Universal Robots URScript: FaiChun_9 Jan_1.script

def Machining1():
  # Default parameters:
  global speed_ms = 0.01
  global speed_rads = 0.75
  global accel_mss = 3
  global accel_radss = 1.2
  global blend_radius_m = 0.0003

  # Add subprograms here
  # Start of main program
  # Program generated by RoboDK v5.6.8 for UR10e on 09/01/2025 14:53:28
  # Using nominal kinematics.
  blend_radius_m = 0.0003
  speed_ms = 0.01
  # set_reference(p[0.305000, -0.155000, 0.000000, 0.000000, 0.000000, 0.000000])
  set_tcp(p[0.000000, 0.000000, 0.252000, 0.000000, 0.000000, 0.000000])
  # Show Tool
  movej([0.378214, -1.028418, -2.649277, -1.034694, 1.570796, 1.949010],accel_radss,speed_rads,0,blend_radius_m)
  movel([0.378214, -1.088062, -2.690368, -0.933959, 1.570796, 1.949010],accel_mss,speed_ms,0,blend_radius_m)
  #SetTool1
  #M_RunCode6
  #SetRPM60000
  speed_ms = 0.01
  #M_RunCode3
  movel([0.378214, -1.116012, -2.706101, -0.890276, 1.570796, 1.949010],accel_mss,speed_ms,0,blend_radius_m)
  speed_ms = 0.003
  movel([0.378214, -1.123422, -2.709978, -0.878989, 1.570796, 1.949010],accel_mss,speed_ms,0,blend_radius_m)
  speed_ms = 0.007
  movel([0.427669, -1.206915, -2.673266, -0.832208, 1.570796, 1.998465],accel_mss,speed_ms,0,blend_radius_m)
  movel([0.418964, -1.213811, -2.669903, -0.828675, 1.570796, 1.989761],accel_mss,speed_ms,0,blend_radius_m)
  movel([0.421470, -1.218334, -2.667668, -0.826387, 1.570796, 1.992267],accel_mss,speed_ms,0,blend_radius_m)
  movel([0.423710, -1.216572, -2.668541, -0.827276, 1.570796, 1.994506],accel_mss,speed_ms,0,blend_radius_m)
  movel([0.422070, -1.213581, -2.670016, -0.828792, 1.570796, 1.992867],accel_mss,speed_ms,0,blend_radius_m)
  movel([0.428515, -1.208497, -2.672499, -0.831392, 1.570796, 1.999312],accel_mss,speed_ms,0,blend_radius_m)
  movel([0.428905, -1.209227, -2.672145, -0.831017, 1.570796, 1.999701],accel_mss,speed_ms,0,blend_radius_m)
  movel([0.430913, -1.212978, -2.670312, -0.829099, 1.570796, 2.001710],accel_mss,speed_ms,0,blend_radius_m)
  movel([0.426574, -1.216377, -2.668637, -0.827374, 1.570796, 1.997371],accel_mss,speed_ms,0,blend_radius_m)
  movel([0.427415, -1.217932, -2.667867, -0.826590, 1.570796, 1.998211],accel_mss,speed_ms,0,blend_radius_m)
  movel([0.431749, -1.214549, -2.669539, -0.828300, 1.570796, 2.002545],accel_mss,speed_ms,0,blend_radius_m)
  movel([0.434110, -1.219016, -2.667329, -0.826045, 1.570796, 2.004906],accel_mss,speed_ms,0,blend_radius_m)
  movel([0.429796, -1.222362, -2.665657, -0.824369, 1.570796, 2.000592],accel_mss,speed_ms,0,blend_radius_m)
  movel([0.431384, -1.225346, -2.664156, -0.822886, 1.570796, 2.002180],accel_mss,speed_ms,0,blend_radius_m)
  movel([0.425058, -1.230240, -2.661672, -0.820476, 1.570796, 1.995855],accel_mss,speed_ms,0,blend_radius_m)
  movel([0.423449, -1.227294, -2.663171, -0.821924, 1.570796, 1.994246],accel_mss,speed_ms,0,blend_radius_m)
  movel([0.421238, -1.229018, -2.662295, -0.821076, 1.570796, 1.992034],accel_mss,speed_ms,0,blend_radius_m)
  movel([0.422852, -1.231953, -2.660796, -0.819639, 1.570796, 1.993648],accel_mss,speed_ms,0,blend_radius_m)
  movel([0.417606, -1.236027, -2.658699, -0.817662, 1.570796, 1.988403],accel_mss,speed_ms,0,blend_radius_m)
  movel([0.416595, -1.236817, -2.658291, -0.817282, 1.570796, 1.987391],accel_mss,speed_ms,0,blend_radius_m)
  movel([0.414170, -1.232527, -2.660502, -0.819360, 1.570796, 1.984966],accel_mss,speed_ms,0,blend_radius_m)
  movel([0.418408, -1.229206, -2.662200, -0.820984, 1.570796, 1.989204],accel_mss,speed_ms,0,blend_radius_m)
  movel([0.417558, -1.227687, -2.662972, -0.821730, 1.570796, 1.988355],accel_mss,speed_ms,0,blend_radius_m)
  movel([0.411120, -1.232746, -2.660390, -0.819253, 1.570796, 1.981917],accel_mss,speed_ms,0,blend_radius_m)
  movel([0.414410, -1.238516, -2.657409, -0.816464, 1.570796, 1.985206],accel_mss,speed_ms,0,blend_radius_m)
  movel([0.308742, -1.323345, -2.608871, -0.780173, 1.570796, 1.879539],accel_mss,speed_ms,0,blend_radius_m)
  movel([0.217512, -1.401117, -2.555954, -0.755318, 1.570796, 1.788308],accel_mss,speed_ms,0,blend_radius_m)
  movel([0.213488, -1.397361, -2.558708, -0.756321, 1.570796, 1.784284],accel_mss,speed_ms,0,blend_radius_m)
  movel([0.208744, -1.401573, -2.555618, -0.755198, 1.570796, 1.779541],accel_mss,speed_ms,0,blend_radius_m)
  movel([0.209793, -1.402537, -2.554907, -0.754944, 1.570796, 1.780589],accel_mss,speed_ms,0,blend_radius_m)
  movel([0.212909, -1.399774, -2.556941, -0.755674, 1.570796, 1.783706],accel_mss,speed_ms,0,blend_radius_m)
  movel([0.215882, -1.402546, -2.554901, -0.754942, 1.570796, 1.786679],accel_mss,speed_ms,0,blend_radius_m)
  movel([0.215131, -1.403208, -2.554412, -0.754769, 1.570796, 1.785928],accel_mss,speed_ms,0,blend_radius_m)
  movel([0.211277, -1.406609, -2.551890, -0.753890, 1.570796, 1.782073],accel_mss,speed_ms,0,blend_radius_m)
  movel([0.209269, -1.404754, -2.553268, -0.754367, 1.570796, 1.780066],accel_mss,speed_ms,0,blend_radius_m)
  movel([0.207663, -1.406180, -2.552209, -0.754000, 1.570796, 1.778459],accel_mss,speed_ms,0,blend_radius_m)
  movel([0.209672, -1.408029, -2.550833, -0.753528, 1.570796, 1.780468],accel_mss,speed_ms,0,blend_radius_m)
  movel([0.205118, -1.412065, -2.547809, -0.752515, 1.570796, 1.775914],accel_mss,speed_ms,0,blend_radius_m)
  movel([0.203102, -1.410238, -2.549181, -0.752970, 1.570796, 1.773898],accel_mss,speed_ms,0,blend_radius_m)
  movel([0.200044, -1.412967, -2.547130, -0.752292, 1.570796, 1.770840],accel_mss,speed_ms,0,blend_radius_m)
  movel([0.197039, -1.410284, -2.549146, -0.752959, 1.570796, 1.767835],accel_mss,speed_ms,0,blend_radius_m)
  movel([0.200101, -1.407535, -2.551201, -0.753653, 1.570796, 1.770897],accel_mss,speed_ms,0,blend_radius_m)
  movel([0.199043, -1.406589, -2.551905, -0.753895, 1.570796, 1.769840],accel_mss,speed_ms,0,blend_radius_m)
  movel([0.195980, -1.409343, -2.549851, -0.753195, 1.570796, 1.766776],accel_mss,speed_ms,0,blend_radius_m)
  movel([0.193434, -1.407104, -2.551522, -0.753763, 1.570796, 1.764230],accel_mss,speed_ms,0,blend_radius_m)
  movel([0.192941, -1.406669, -2.551845, -0.753874, 1.570796, 1.763737],accel_mss,speed_ms,0,blend_radius_m)
  movel([0.197491, -1.402558, -2.554892, -0.754939, 1.570796, 1.768287],accel_mss,speed_ms,0,blend_radius_m)
  movel([0.199540, -1.404383, -2.553543, -0.754463, 1.570796, 1.770337],accel_mss,speed_ms,0,blend_radius_m)
  movel([0.201142, -1.402944, -2.554607, -0.754838, 1.570796, 1.771938],accel_mss,speed_ms,0,blend_radius_m)
  movel([0.198026, -1.400161, -2.556657, -0.755571, 1.570796, 1.768823],accel_mss,speed_ms,0,blend_radius_m)
  movel([0.191871, -1.405733, -2.552541, -0.754115, 1.570796, 1.762667],accel_mss,speed_ms,0,blend_radius_m)
  movel([0.191373, -1.405301, -2.552862, -0.754226, 1.570796, 1.762169],accel_mss,speed_ms,0,blend_radius_m)
  movel([0.131815, -1.358213, -2.586196, -0.767981, 1.570796, 1.702611],accel_mss,speed_ms,0,blend_radius_m)
  movel([0.062823, -1.314529, -2.614344, -0.783517, 1.570796, 1.633619],accel_mss,speed_ms,0,blend_radius_m)
  movel([0.069044, -1.307429, -2.618676, -0.786284, 1.570796, 1.639841],accel_mss,speed_ms,0,blend_radius_m)
  movel([0.064886, -1.305093, -2.620087, -0.787209, 1.570796, 1.635683],accel_mss,speed_ms,0,blend_radius_m)
  movel([0.063265, -1.306951, -2.618965, -0.786472, 1.570796, 1.634061],accel_mss,speed_ms,0,blend_radius_m)
  movel([0.066004, -1.308479, -2.618039, -0.785870, 1.570796, 1.636801],accel_mss,speed_ms,0,blend_radius_m)
  movel([0.061405, -1.313734, -2.614831, -0.783823, 1.570796, 1.632201],accel_mss,speed_ms,0,blend_radius_m)
  movel([0.060750, -1.313370, -2.615055, -0.783964, 1.570796, 1.631546],accel_mss,speed_ms,0,blend_radius_m)
  movel([0.057348, -1.311503, -2.616198, -0.784688, 1.570796, 1.628144],accel_mss,speed_ms,0,blend_radius_m)
  movel([0.060443, -1.307941, -2.618366, -0.786082, 1.570796, 1.631240],accel_mss,speed_ms,0,blend_radius_m)
  movel([0.059013, -1.307156, -2.618841, -0.786392, 1.570796, 1.629809],accel_mss,speed_ms,0,blend_radius_m)
  movel([0.055918, -1.310726, -2.616672, -0.784991, 1.570796, 1.626714],accel_mss,speed_ms,0,blend_radius_m)
  movel([0.051821, -1.308523, -2.618013, -0.785853, 1.570796, 1.622617],accel_mss,speed_ms,0,blend_radius_m)
  movel([0.054912, -1.304932, -2.620184, -0.787273, 1.570796, 1.625709],accel_mss,speed_ms,0,blend_radius_m)
  movel([0.052126, -1.303438, -2.621082, -0.787868, 1.570796, 1.622923],accel_mss,speed_ms,0,blend_radius_m)
  movel([0.056741, -1.298064, -2.624290, -0.790035, 1.570796, 1.627538],accel_mss,speed_ms,0,blend_radius_m)
  movel([0.059531, -1.299576, -2.623391, -0.789421, 1.570796, 1.630327],accel_mss,speed_ms,0,blend_radius_m)
  movel([0.061161, -1.297689, -2.624513, -0.790187, 1.570796, 1.631957],accel_mss,speed_ms,0,blend_radius_m)
  movel([0.058371, -1.296169, -2.625412, -0.790807, 1.570796, 1.629167],accel_mss,speed_ms,0,blend_radius_m)
  movel([0.062287, -1.291620, -2.628088, -0.792681, 1.570796, 1.633084],accel_mss,speed_ms,0,blend_radius_m)
  movel([0.063052, -1.290735, -2.628605, -0.793049, 1.570796, 1.633848],accel_mss,speed_ms,0,blend_radius_m)
  movel([0.067186, -1.293020, -2.627267, -0.792102, 1.570796, 1.637983],accel_mss,speed_ms,0,blend_radius_m)
  movel([0.064017, -1.296673, -2.625115, -0.790602, 1.570796, 1.634813],accel_mss,speed_ms,0,blend_radius_m)
  movel([0.065457, -1.297471, -2.624642, -0.790276, 1.570796, 1.636253],accel_mss,speed_ms,0,blend_radius_m)
  movel([0.070282, -1.291926, -2.627908, -0.792554, 1.570796, 1.641079],accel_mss,speed_ms,0,blend_radius_m)
  movel([0.064708, -1.288816, -2.629723, -0.793850, 1.570796, 1.635504],accel_mss,speed_ms,0,blend_radius_m)
  movel([0.160316, -1.180338, -2.685740, -0.846311, 1.570796, 1.731113],accel_mss,speed_ms,0,blend_radius_m)
  movel([0.277315, -1.052375, -2.735928, -0.924086, 1.570796, 1.848111],accel_mss,speed_ms,0,blend_radius_m)
  movel([0.278486, -1.051118, -2.736347, -0.924924, 1.570796, 1.849282],accel_mss,speed_ms,0,blend_radius_m)
  movel([0.283865, -1.056777, -2.734448, -0.921164, 1.570796, 1.854661],accel_mss,speed_ms,0,blend_radius_m)
  movel([0.291287, -1.048884, -2.737089, -0.926415, 1.570796, 1.862083],accel_mss,speed_ms,0,blend_radius_m)
  movel([0.289909, -1.047384, -2.737586, -0.927419, 1.570796, 1.860706],accel_mss,speed_ms,0,blend_radius_m)
  movel([0.285009, -1.052605, -2.735851, -0.923933, 1.570796, 1.855805],accel_mss,speed_ms,0,blend_radius_m)
  movel([0.281034, -1.048391, -2.737253, -0.926745, 1.570796, 1.851830],accel_mss,speed_ms,0,blend_radius_m)
  movel([0.282209, -1.047128, -2.737670, -0.927591, 1.570796, 1.853005],accel_mss,speed_ms,0,blend_radius_m)
  movel([0.288325, -1.040563, -2.739819, -0.932008, 1.570796, 1.859122],accel_mss,speed_ms,0,blend_radius_m)
  movel([0.291001, -1.043464, -2.738874, -0.930052, 1.570796, 1.861797],accel_mss,speed_ms,0,blend_radius_m)
  movel([0.293574, -1.040720, -2.739767, -0.931902, 1.570796, 1.864371],accel_mss,speed_ms,0,blend_radius_m)
  movel([0.290903, -1.037800, -2.740712, -0.933877, 1.570796, 1.861699],accel_mss,speed_ms,0,blend_radius_m)
  movel([0.298320, -1.029861, -2.743245, -0.939282, 1.570796, 1.869116],accel_mss,speed_ms,0,blend_radius_m)
  movel([0.300982, -1.032832, -2.742303, -0.937254, 1.570796, 1.871778],accel_mss,speed_ms,0,blend_radius_m)
  movel([0.306035, -1.027460, -2.744002, -0.940927, 1.570796, 1.876831],accel_mss,speed_ms,0,blend_radius_m)
  movel([0.309920, -1.031931, -2.742590, -0.937868, 1.570796, 1.880716],accel_mss,speed_ms,0,blend_radius_m)
  movel([0.304877, -1.037251, -2.740889, -0.934249, 1.570796, 1.875674],accel_mss,speed_ms,0,blend_radius_m)
  movel([0.306232, -1.038803, -2.740388, -0.933198, 1.570796, 1.877028],accel_mss,speed_ms,0,blend_radius_m)
  movel([0.311270, -1.033502, -2.742090, -0.936797, 1.570796, 1.882066],accel_mss,speed_ms,0,blend_radius_m)
  movel([0.315085, -1.038000, -2.740648, -0.933742, 1.570796, 1.885882],accel_mss,speed_ms,0,blend_radius_m)
  movel([0.307670, -1.045746, -2.738125, -0.928518, 1.570796, 1.878466],accel_mss,speed_ms,0,blend_radius_m)
  movel([0.305079, -1.042766, -2.739101, -0.930521, 1.570796, 1.875875],accel_mss,speed_ms,0,blend_radius_m)
  movel([0.302496, -1.045482, -2.738212, -0.928695, 1.570796, 1.873292],accel_mss,speed_ms,0,blend_radius_m)
  movel([0.306428, -1.049986, -2.736724, -0.925679, 1.570796, 1.877224],accel_mss,speed_ms,0,blend_radius_m)
  movel([0.316412, -1.039578, -2.740138, -0.932673, 1.570796, 1.887209],accel_mss,speed_ms,0,blend_radius_m)
  movel([0.378214, -1.123422, -2.709978, -0.878989, 1.570796, 1.949010],accel_mss,speed_ms,0,blend_radius_m)
  speed_ms = 0.003
  movel([0.378214, -1.116012, -2.706101, -0.890276, 1.570796, 1.949010],accel_mss,speed_ms,0,blend_radius_m)
  speed_ms = 1.000
  movel([0.378214, -1.088062, -2.690368, -0.933959, 1.570796, 1.949010],accel_mss,speed_ms,0,blend_radius_m)
  #M_RunCode9
  movel([0.299608, -1.056483, -2.701958, -0.953949, 1.570796, 1.870404],accel_mss,speed_ms,0,blend_radius_m)
  #M_RunCode3
  movel([0.299608, -1.084408, -2.718093, -0.909888, 1.570796, 1.870404],accel_mss,speed_ms,0,blend_radius_m)
  speed_ms = 0.003
  movel([0.299608, -1.091834, -2.722073, -0.898483, 1.570796, 1.870404],accel_mss,speed_ms,0,blend_radius_m)
  speed_ms = 0.007
  movel([0.297554, -1.094394, -2.721127, -0.896868, 1.570796, 1.868350],accel_mss,speed_ms,0,blend_radius_m)
  movel([0.295269, -1.096439, -2.720366, -0.895583, 1.570796, 1.866066],accel_mss,speed_ms,0,blend_radius_m)
  movel([0.292750, -1.097981, -2.719791, -0.894617, 1.570796, 1.863546],accel_mss,speed_ms,0,blend_radius_m)
  movel([0.289989, -1.099020, -2.719402, -0.893967, 1.570796, 1.860786],accel_mss,speed_ms,0,blend_radius_m)
  movel([0.287614, -1.099423, -2.719251, -0.893715, 1.570796, 1.858411],accel_mss,speed_ms,0,blend_radius_m)
  movel([0.285561, -1.099227, -2.719324, -0.893838, 1.570796, 1.856357],accel_mss,speed_ms,0,blend_radius_m)
  movel([0.283804, -1.098580, -2.719567, -0.894242, 1.570796, 1.854601],accel_mss,speed_ms,0,blend_radius_m)
  movel([0.282319, -1.097620, -2.719926, -0.894843, 1.570796, 1.853116],accel_mss,speed_ms,0,blend_radius_m)
  movel([0.279271, -1.094519, -2.721080, -0.896790, 1.570796, 1.850068],accel_mss,speed_ms,0,blend_radius_m)
  movel([0.276341, -1.091631, -2.722147, -0.898610, 1.570796, 1.847137],accel_mss,speed_ms,0,blend_radius_m)
  movel([0.274975, -1.090758, -2.722469, -0.899163, 1.570796, 1.845772],accel_mss,speed_ms,0,blend_radius_m)
  movel([0.273381, -1.090179, -2.722681, -0.899529, 1.570796, 1.844178],accel_mss,speed_ms,0,blend_radius_m)
  movel([0.271551, -1.090019, -2.722740, -0.899630, 1.570796, 1.842347],accel_mss,speed_ms,0,blend_radius_m)
  movel([0.269474, -1.090407, -2.722597, -0.899385, 1.570796, 1.840271],accel_mss,speed_ms,0,blend_radius_m)
  movel([0.269162, -1.091589, -2.722163, -0.898637, 1.570796, 1.839958],accel_mss,speed_ms,0,blend_radius_m)
  movel([0.268451, -1.094807, -2.720973, -0.896608, 1.570796, 1.839247],accel_mss,speed_ms,0,blend_radius_m)
  movel([0.268160, -1.097519, -2.719963, -0.894906, 1.570796, 1.838957],accel_mss,speed_ms,0,blend_radius_m)
  movel([0.268285, -1.099732, -2.719135, -0.893522, 1.570796, 1.839081],accel_mss,speed_ms,0,blend_radius_m)
  movel([0.268822, -1.101454, -2.718487, -0.892448, 1.570796, 1.839618],accel_mss,speed_ms,0,blend_radius_m)
  movel([0.269704, -1.102726, -2.718006, -0.891657, 1.570796, 1.840500],accel_mss,speed_ms,0,blend_radius_m)
  movel([0.270877, -1.103589, -2.717679, -0.891120, 1.570796, 1.841674],accel_mss,speed_ms,0,blend_radius_m)
  movel([0.272340, -1.104040, -2.717508, -0.890841, 1.570796, 1.843137],accel_mss,speed_ms,0,blend_radius_m)
  movel([0.274092, -1.104087, -2.717491, -0.890812, 1.570796, 1.844889],accel_mss,speed_ms,0,blend_radius_m)
  movel([0.264197, -1.106964, -2.716395, -0.889030, 1.570796, 1.834993],accel_mss,speed_ms,0,blend_radius_m)
  movel([0.272508, -1.075450, -2.727989, -0.908949, 1.570796, 1.843305],accel_mss,speed_ms,0,blend_radius_m)
  movel([0.273532, -1.075136, -2.728101, -0.909153, 1.570796, 1.844329],accel_mss,speed_ms,0,blend_radius_m)
  movel([0.276027, -1.074709, -2.728251, -0.909429, 1.570796, 1.846823],accel_mss,speed_ms,0,blend_radius_m)
  movel([0.278273, -1.075047, -2.728132, -0.909210, 1.570796, 1.849069],accel_mss,speed_ms,0,blend_radius_m)
  movel([0.280254, -1.075949, -2.727812, -0.908627, 1.570796, 1.851051],accel_mss,speed_ms,0,blend_radius_m)
  movel([0.281955, -1.077216, -2.727363, -0.907810, 1.570796, 1.852751],accel_mss,speed_ms,0,blend_radius_m)
  movel([0.285849, -1.081361, -2.725882, -0.905146, 1.570796, 1.856646],accel_mss,speed_ms,0,blend_radius_m)
  movel([0.289358, -1.085288, -2.724465, -0.902636, 1.570796, 1.860155],accel_mss,speed_ms,0,blend_radius_m)
  movel([0.290895, -1.086507, -2.724022, -0.901859, 1.570796, 1.861691],accel_mss,speed_ms,0,blend_radius_m)
  movel([0.292636, -1.087385, -2.723703, -0.901301, 1.570796, 1.863432],accel_mss,speed_ms,0,blend_radius_m)
  movel([0.294569, -1.087761, -2.723566, -0.901062, 1.570796, 1.865365],accel_mss,speed_ms,0,blend_radius_m)
  movel([0.296672, -1.087485, -2.723667, -0.901238, 1.570796, 1.867469],accel_mss,speed_ms,0,blend_radius_m)
  movel([0.299389, -1.086337, -2.724084, -0.901968, 1.570796, 1.870185],accel_mss,speed_ms,0,blend_radius_m)
  movel([0.300577, -1.085516, -2.724383, -0.902491, 1.570796, 1.871373],accel_mss,speed_ms,0,blend_radius_m)
  movel([0.301654, -1.084522, -2.724743, -0.903125, 1.570796, 1.872450],accel_mss,speed_ms,0,blend_radius_m)
  movel([0.303363, -1.082314, -2.725539, -0.904535, 1.570796, 1.874159],accel_mss,speed_ms,0,blend_radius_m)
  movel([0.304392, -1.080010, -2.726366, -0.906013, 1.570796, 1.875188],accel_mss,speed_ms,0,blend_radius_m)
  movel([0.304681, -1.078561, -2.726884, -0.906944, 1.570796, 1.875477],accel_mss,speed_ms,0,blend_radius_m)
  movel([0.304556, -1.077581, -2.727233, -0.907575, 1.570796, 1.875352],accel_mss,speed_ms,0,blend_radius_m)
  movel([0.304086, -1.077081, -2.727411, -0.907897, 1.570796, 1.874882],accel_mss,speed_ms,0,blend_radius_m)
  movel([0.303340, -1.077079, -2.727412, -0.907898, 1.570796, 1.874137],accel_mss,speed_ms,0,blend_radius_m)
  movel([0.301979, -1.077952, -2.727101, -0.907336, 1.570796, 1.872776],accel_mss,speed_ms,0,blend_radius_m)
  movel([0.300659, -1.078907, -2.726761, -0.906722, 1.570796, 1.871455],accel_mss,speed_ms,0,blend_radius_m)
  movel([0.299075, -1.079565, -2.726526, -0.906298, 1.570796, 1.869871],accel_mss,speed_ms,0,blend_radius_m)
  movel([0.297392, -1.079689, -2.726481, -0.906219, 1.570796, 1.868188],accel_mss,speed_ms,0,blend_radius_m)
  movel([0.296382, -1.078930, -2.726752, -0.906706, 1.570796, 1.867179],accel_mss,speed_ms,0,blend_radius_m)
  movel([0.296029, -1.077505, -2.727260, -0.907624, 1.570796, 1.866825],accel_mss,speed_ms,0,blend_radius_m)
  movel([0.296310, -1.075635, -2.727924, -0.908830, 1.570796, 1.867107],accel_mss,speed_ms,0,blend_radius_m)
  movel([0.297148, -1.073602, -2.728642, -0.910145, 1.570796, 1.867945],accel_mss,speed_ms,0,blend_radius_m)
  movel([0.298463, -1.071693, -2.729313, -0.911383, 1.570796, 1.869259],accel_mss,speed_ms,0,blend_radius_m)
  movel([0.300143, -1.070159, -2.729850, -0.912380, 1.570796, 1.870939],accel_mss,speed_ms,0,blend_radius_m)
  movel([0.302063, -1.069262, -2.730163, -0.912964, 1.570796, 1.872860],accel_mss,speed_ms,0,blend_radius_m)
  movel([0.303592, -1.069033, -2.730242, -0.913113, 1.570796, 1.874388],accel_mss,speed_ms,0,blend_radius_m)
  movel([0.304794, -1.069305, -2.730148, -0.912936, 1.570796, 1.875590],accel_mss,speed_ms,0,blend_radius_m)
  movel([0.305666, -1.070083, -2.729876, -0.912430, 1.570796, 1.876463],accel_mss,speed_ms,0,blend_radius_m)
  movel([0.306212, -1.071354, -2.729432, -0.911603, 1.570796, 1.877008],accel_mss,speed_ms,0,blend_radius_m)
  movel([0.306451, -1.073019, -2.728847, -0.910523, 1.570796, 1.877247],accel_mss,speed_ms,0,blend_radius_m)
  movel([0.306392, -1.074975, -2.728157, -0.909257, 1.570796, 1.877188],accel_mss,speed_ms,0,blend_radius_m)
  movel([0.305401, -1.079734, -2.726465, -0.906190, 1.570796, 1.876198],accel_mss,speed_ms,0,blend_radius_m)
  movel([0.304321, -1.082915, -2.725323, -0.904151, 1.570796, 1.875117],accel_mss,speed_ms,0,blend_radius_m)
  movel([0.302996, -1.085992, -2.724210, -0.902187, 1.570796, 1.873793],accel_mss,speed_ms,0,blend_radius_m)
  movel([0.301425, -1.088961, -2.723127, -0.900301, 1.570796, 1.872221],accel_mss,speed_ms,0,blend_radius_m)
  movel([0.299608, -1.091834, -2.722073, -0.898483, 1.570796, 1.870404],accel_mss,speed_ms,0,blend_radius_m)
  speed_ms = 0.003
  movel([0.299608, -1.084408, -2.718093, -0.909888, 1.570796, 1.870404],accel_mss,speed_ms,0,blend_radius_m)
  speed_ms = 1.000
  movel([0.299608, -1.056483, -2.701958, -0.953949, 1.570796, 1.870404],accel_mss,speed_ms,0,blend_radius_m)
  #M_RunCode9
  movel([0.290804, -1.078007, -2.694153, -0.940229, 1.570796, 1.861601],accel_mss,speed_ms,0,blend_radius_m)
  #M_RunCode3
  movel([0.290804, -1.105959, -2.710015, -0.896415, 1.570796, 1.861601],accel_mss,speed_ms,0,blend_radius_m)
  speed_ms = 0.003
  movel([0.290804, -1.113377, -2.713924, -0.885087, 1.570796, 1.861601],accel_mss,speed_ms,0,blend_radius_m)
  speed_ms = 0.007
  movel([0.292487, -1.113483, -2.713883, -0.885022, 1.570796, 1.863283],accel_mss,speed_ms,0,blend_radius_m)
  movel([0.293570, -1.113959, -2.713698, -0.884731, 1.570796, 1.864366],accel_mss,speed_ms,0,blend_radius_m)
  movel([0.294059, -1.114807, -2.713368, -0.884213, 1.570796, 1.864855],accel_mss,speed_ms,0,blend_radius_m)
  movel([0.293950, -1.116023, -2.712894, -0.883472, 1.570796, 1.864746],accel_mss,speed_ms,0,blend_radius_m)
  movel([0.293317, -1.117375, -2.712365, -0.882649, 1.570796, 1.864113],accel_mss,speed_ms,0,blend_radius_m)
  movel([0.292224, -1.118630, -2.711872, -0.881887, 1.570796, 1.863020],accel_mss,speed_ms,0,blend_radius_m)
  movel([0.290678, -1.119787, -2.711417, -0.881185, 1.570796, 1.861474],accel_mss,speed_ms,0,blend_radius_m)
  movel([0.288670, -1.120856, -2.710995, -0.880538, 1.570796, 1.859466],accel_mss,speed_ms,0,blend_radius_m)
  movel([0.283159, -1.122966, -2.710159, -0.879264, 1.570796, 1.853956],accel_mss,speed_ms,0,blend_radius_m)
  movel([0.275572, -1.125220, -2.709261, -0.877908, 1.570796, 1.846369],accel_mss,speed_ms,0,blend_radius_m)
  movel([0.268111, -1.127055, -2.708527, -0.876807, 1.570796, 1.838907],accel_mss,speed_ms,0,blend_radius_m)
  movel([0.262988, -1.127840, -2.708211, -0.876337, 1.570796, 1.833785],accel_mss,speed_ms,0,blend_radius_m)
  movel([0.261301, -1.127782, -2.708235, -0.876372, 1.570796, 1.832097],accel_mss,speed_ms,0,blend_radius_m)
  movel([0.260198, -1.127357, -2.708406, -0.876627, 1.570796, 1.830994],accel_mss,speed_ms,0,blend_radius_m)
  movel([0.259674, -1.126556, -2.708727, -0.877106, 1.570796, 1.830471],accel_mss,speed_ms,0,blend_radius_m)
  movel([0.259738, -1.125376, -2.709199, -0.877814, 1.570796, 1.830535],accel_mss,speed_ms,0,blend_radius_m)
  movel([0.260326, -1.124046, -2.709729, -0.878613, 1.570796, 1.831122],accel_mss,speed_ms,0,blend_radius_m)
  movel([0.261388, -1.122787, -2.710230, -0.879372, 1.570796, 1.832184],accel_mss,speed_ms,0,blend_radius_m)
  movel([0.262917, -1.121604, -2.710699, -0.880086, 1.570796, 1.833713],accel_mss,speed_ms,0,blend_radius_m)
  movel([0.264922, -1.120492, -2.711139, -0.880758, 1.570796, 1.835718],accel_mss,speed_ms,0,blend_radius_m)
  movel([0.270463, -1.118269, -2.712014, -0.882106, 1.570796, 1.841260],accel_mss,speed_ms,0,blend_radius_m)
  movel([0.278124, -1.115921, -2.712934, -0.883534, 1.570796, 1.848920],accel_mss,speed_ms,0,blend_radius_m)
  movel([0.285652, -1.114089, -2.713648, -0.884652, 1.570796, 1.856449],accel_mss,speed_ms,0,blend_radius_m)
  movel([0.290804, -1.113377, -2.713924, -0.885087, 1.570796, 1.861601],accel_mss,speed_ms,0,blend_radius_m)
  speed_ms = 0.003
  movel([0.290804, -1.105959, -2.710015, -0.896415, 1.570796, 1.861601],accel_mss,speed_ms,0,blend_radius_m)
  speed_ms = 1.000
  movel([0.290804, -1.078007, -2.694153, -0.940229, 1.570796, 1.861601],accel_mss,speed_ms,0,blend_radius_m)
  #M_RunCode9
  movel([0.295393, -1.074864, -2.695318, -0.942207, 1.570796, 1.866190],accel_mss,speed_ms,0,blend_radius_m)
  #M_RunCode3
  movel([0.295393, -1.102816, -2.711220, -0.898354, 1.570796, 1.866190],accel_mss,speed_ms,0,blend_radius_m)
  speed_ms = 0.003
  movel([0.295393, -1.110235, -2.715139, -0.887014, 1.570796, 1.866190],accel_mss,speed_ms,0,blend_radius_m)
  speed_ms = 0.007
  movel([0.295505, -1.111918, -2.714490, -0.885981, 1.570796, 1.866301],accel_mss,speed_ms,0,blend_radius_m)
  movel([0.295326, -1.113772, -2.713771, -0.884846, 1.570796, 1.866122],accel_mss,speed_ms,0,blend_radius_m)
  movel([0.294860, -1.115787, -2.712986, -0.883616, 1.570796, 1.865656],accel_mss,speed_ms,0,blend_radius_m)
  movel([0.294140, -1.117864, -2.712173, -0.882351, 1.570796, 1.864936],accel_mss,speed_ms,0,blend_radius_m)
  movel([0.293196, -1.119900, -2.711373, -0.881117, 1.570796, 1.863992],accel_mss,speed_ms,0,blend_radius_m)
  movel([0.292028, -1.121889, -2.710586, -0.879914, 1.570796, 1.862824],accel_mss,speed_ms,0,blend_radius_m)
  movel([0.290637, -1.123836, -2.709813, -0.878740, 1.570796, 1.861434],accel_mss,speed_ms,0,blend_radius_m)
  movel([0.289037, -1.125708, -2.709066, -0.877615, 1.570796, 1.859834],accel_mss,speed_ms,0,blend_radius_m)
  movel([0.287243, -1.127464, -2.708362, -0.876562, 1.570796, 1.858040],accel_mss,speed_ms,0,blend_radius_m)
  movel([0.285249, -1.129114, -2.707699, -0.875576, 1.570796, 1.856046],accel_mss,speed_ms,0,blend_radius_m)
  movel([0.283057, -1.130656, -2.707076, -0.874657, 1.570796, 1.853853],accel_mss,speed_ms,0,blend_radius_m)
  movel([0.280704, -1.132048, -2.706511, -0.873829, 1.570796, 1.851500],accel_mss,speed_ms,0,blend_radius_m)
  movel([0.278220, -1.133257, -2.706020, -0.873112, 1.570796, 1.849017],accel_mss,speed_ms,0,blend_radius_m)
  movel([0.275609, -1.134281, -2.705602, -0.872505, 1.570796, 1.846406],accel_mss,speed_ms,0,blend_radius_m)
  movel([0.272869, -1.135123, -2.705259, -0.872007, 1.570796, 1.843665],accel_mss,speed_ms,0,blend_radius_m)
  movel([0.270190, -1.135733, -2.705009, -0.871647, 1.570796, 1.840986],accel_mss,speed_ms,0,blend_radius_m)
  movel([0.267774, -1.136056, -2.704876, -0.871456, 1.570796, 1.838571],accel_mss,speed_ms,0,blend_radius_m)
  movel([0.265617, -1.136094, -2.704861, -0.871434, 1.570796, 1.836414],accel_mss,speed_ms,0,blend_radius_m)
  movel([0.263719, -1.135848, -2.704962, -0.871579, 1.570796, 1.834516],accel_mss,speed_ms,0,blend_radius_m)
  movel([0.262095, -1.135340, -2.705170, -0.871879, 1.570796, 1.832892],accel_mss,speed_ms,0,blend_radius_m)
  movel([0.260758, -1.134598, -2.705473, -0.872318, 1.570796, 1.831554],accel_mss,speed_ms,0,blend_radius_m)
  movel([0.259709, -1.133623, -2.705871, -0.872895, 1.570796, 1.830505],accel_mss,speed_ms,0,blend_radius_m)
  movel([0.258949, -1.132408, -2.706365, -0.873616, 1.570796, 1.829745],accel_mss,speed_ms,0,blend_radius_m)
  movel([0.258474, -1.130987, -2.706942, -0.874460, 1.570796, 1.829271],accel_mss,speed_ms,0,blend_radius_m)
  movel([0.258285, -1.129391, -2.707587, -0.875411, 1.570796, 1.829081],accel_mss,speed_ms,0,blend_radius_m)
  movel([0.258385, -1.127612, -2.708303, -0.876474, 1.570796, 1.829181],accel_mss,speed_ms,0,blend_radius_m)
  movel([0.258770, -1.125654, -2.709088, -0.877647, 1.570796, 1.829567],accel_mss,speed_ms,0,blend_radius_m)
  movel([0.259418, -1.123617, -2.709900, -0.878872, 1.570796, 1.830215],accel_mss,speed_ms,0,blend_radius_m)
  movel([0.260304, -1.121597, -2.710702, -0.880090, 1.570796, 1.831100],accel_mss,speed_ms,0,blend_radius_m)
  movel([0.261431, -1.119598, -2.711491, -0.881299, 1.570796, 1.832228],accel_mss,speed_ms,0,blend_radius_m)
  movel([0.262801, -1.117618, -2.712270, -0.882501, 1.570796, 1.833597],accel_mss,speed_ms,0,blend_radius_m)
  movel([0.264397, -1.115694, -2.713023, -0.883673, 1.570796, 1.835194],accel_mss,speed_ms,0,blend_radius_m)
  movel([0.266204, -1.113865, -2.713735, -0.884789, 1.570796, 1.837001],accel_mss,speed_ms,0,blend_radius_m)
  movel([0.268225, -1.112137, -2.714405, -0.885847, 1.570796, 1.839021],accel_mss,speed_ms,0,blend_radius_m)
  movel([0.270457, -1.110505, -2.715036, -0.886849, 1.570796, 1.841253],accel_mss,speed_ms,0,blend_radius_m)
  movel([0.272869, -1.109019, -2.715608, -0.887763, 1.570796, 1.843665],accel_mss,speed_ms,0,blend_radius_m)
  movel([0.275418, -1.107721, -2.716105, -0.888563, 1.570796, 1.846215],accel_mss,speed_ms,0,blend_radius_m)
  movel([0.278109, -1.106616, -2.716528, -0.889245, 1.570796, 1.848905],accel_mss,speed_ms,0,blend_radius_m)
  movel([0.280939, -1.105707, -2.716874, -0.889807, 1.570796, 1.851735],accel_mss,speed_ms,0,blend_radius_m)
  movel([0.283697, -1.105056, -2.717122, -0.890211, 1.570796, 1.854493],accel_mss,speed_ms,0,blend_radius_m)
  movel([0.286181, -1.104717, -2.717251, -0.890421, 1.570796, 1.856977],accel_mss,speed_ms,0,blend_radius_m)
  movel([0.288389, -1.104690, -2.717261, -0.890437, 1.570796, 1.859186],accel_mss,speed_ms,0,blend_radius_m)
  movel([0.290319, -1.104973, -2.717154, -0.890262, 1.570796, 1.861115],accel_mss,speed_ms,0,blend_radius_m)
  movel([0.291955, -1.105538, -2.716939, -0.889912, 1.570796, 1.862751],accel_mss,speed_ms,0,blend_radius_m)
  movel([0.293278, -1.106350, -2.716629, -0.889410, 1.570796, 1.864075],accel_mss,speed_ms,0,blend_radius_m)
  movel([0.294289, -1.107413, -2.716223, -0.888753, 1.570796, 1.865085],accel_mss,speed_ms,0,blend_radius_m)
  movel([0.294991, -1.108722, -2.715721, -0.887946, 1.570796, 1.865787],accel_mss,speed_ms,0,blend_radius_m)
  movel([0.295393, -1.110235, -2.715139, -0.887014, 1.570796, 1.866190],accel_mss,speed_ms,0,blend_radius_m)
  speed_ms = 0.003
  movel([0.295393, -1.102816, -2.711220, -0.898354, 1.570796, 1.866190],accel_mss,speed_ms,0,blend_radius_m)
  speed_ms = 1.000
  movel([0.295393, -1.074864, -2.695318, -0.942207, 1.570796, 1.866190],accel_mss,speed_ms,0,blend_radius_m)
  #M_RunCode9
  movel([0.205944, -1.317083, -2.576173, -0.819133, 1.570796, 1.776740],accel_mss,speed_ms,0,blend_radius_m)
  #M_RunCode3
  movel([0.205944, -1.342817, -2.588898, -0.780673, 1.570796, 1.776740],accel_mss,speed_ms,0,blend_radius_m)
  speed_ms = 0.003
  movel([0.205944, -1.349516, -2.592008, -0.770866, 1.570796, 1.776740],accel_mss,speed_ms,0,blend_radius_m)
  speed_ms = 0.007
  movel([0.207811, -1.349362, -2.592110, -0.770918, 1.570796, 1.778607],accel_mss,speed_ms,0,blend_radius_m)
  movel([0.209531, -1.349695, -2.591889, -0.770805, 1.570796, 1.780327],accel_mss,speed_ms,0,blend_radius_m)
  movel([0.211081, -1.350383, -2.591433, -0.770573, 1.570796, 1.781877],accel_mss,speed_ms,0,blend_radius_m)
  movel([0.212441, -1.351297, -2.590826, -0.770266, 1.570796, 1.783238],accel_mss,speed_ms,0,blend_radius_m)
  movel([0.215631, -1.354207, -2.588886, -0.769296, 1.570796, 1.786427],accel_mss,speed_ms,0,blend_radius_m)
  movel([0.218525, -1.356949, -2.587046, -0.768393, 1.570796, 1.789322],accel_mss,speed_ms,0,blend_radius_m)
  movel([0.219761, -1.357825, -2.586457, -0.768107, 1.570796, 1.790557],accel_mss,speed_ms,0,blend_radius_m)
  movel([0.221138, -1.358481, -2.586015, -0.767893, 1.570796, 1.791935],accel_mss,speed_ms,0,blend_radius_m)
  movel([0.222629, -1.358814, -2.585790, -0.767785, 1.570796, 1.793425],accel_mss,speed_ms,0,blend_radius_m)
  movel([0.224213, -1.358726, -2.585850, -0.767814, 1.570796, 1.795009],accel_mss,speed_ms,0,blend_radius_m)
  movel([0.226211, -1.358094, -2.586275, -0.768019, 1.570796, 1.797008],accel_mss,speed_ms,0,blend_radius_m)
  movel([0.227066, -1.357605, -2.586605, -0.768179, 1.570796, 1.797862],accel_mss,speed_ms,0,blend_radius_m)
  movel([0.227828, -1.357000, -2.587013, -0.768377, 1.570796, 1.798625],accel_mss,speed_ms,0,blend_radius_m)
  movel([0.228991, -1.355630, -2.587932, -0.768826, 1.570796, 1.799788],accel_mss,speed_ms,0,blend_radius_m)
  movel([0.229636, -1.354166, -2.588913, -0.769310, 1.570796, 1.800433],accel_mss,speed_ms,0,blend_radius_m)
  movel([0.229767, -1.353231, -2.589538, -0.769620, 1.570796, 1.800564],accel_mss,speed_ms,0,blend_radius_m)
  movel([0.229613, -1.352583, -2.589970, -0.769836, 1.570796, 1.800410],accel_mss,speed_ms,0,blend_radius_m)
  movel([0.229225, -1.352237, -2.590200, -0.769952, 1.570796, 1.800022],accel_mss,speed_ms,0,blend_radius_m)
  movel([0.228657, -1.352201, -2.590224, -0.769964, 1.570796, 1.799454],accel_mss,speed_ms,0,blend_radius_m)
  movel([0.227679, -1.352710, -2.589885, -0.769794, 1.570796, 1.798476],accel_mss,speed_ms,0,blend_radius_m)
  movel([0.226731, -1.353276, -2.589507, -0.769605, 1.570796, 1.797528],accel_mss,speed_ms,0,blend_radius_m)
  movel([0.225568, -1.353636, -2.589267, -0.769486, 1.570796, 1.796364],accel_mss,speed_ms,0,blend_radius_m)
  movel([0.224298, -1.353642, -2.589263, -0.769484, 1.570796, 1.795094],accel_mss,speed_ms,0,blend_radius_m)
  movel([0.223489, -1.353098, -2.589626, -0.769665, 1.570796, 1.794285],accel_mss,speed_ms,0,blend_radius_m)
  movel([0.223135, -1.352151, -2.590258, -0.769980, 1.570796, 1.793932],accel_mss,speed_ms,0,blend_radius_m)
  movel([0.223236, -1.350938, -2.591064, -0.770386, 1.570796, 1.794032],accel_mss,speed_ms,0,blend_radius_m)
  movel([0.223753, -1.349647, -2.591921, -0.770821, 1.570796, 1.794549],accel_mss,speed_ms,0,blend_radius_m)
  movel([0.224636, -1.348461, -2.592705, -0.771222, 1.570796, 1.795432],accel_mss,speed_ms,0,blend_radius_m)
  movel([0.225814, -1.347538, -2.593315, -0.771536, 1.570796, 1.796610],accel_mss,speed_ms,0,blend_radius_m)
  movel([0.227215, -1.347042, -2.593642, -0.771705, 1.570796, 1.798012],accel_mss,speed_ms,0,blend_radius_m)
  movel([0.228360, -1.346963, -2.593694, -0.771732, 1.570796, 1.799156],accel_mss,speed_ms,0,blend_radius_m)
  movel([0.229286, -1.347196, -2.593540, -0.771653, 1.570796, 1.800083],accel_mss,speed_ms,0,blend_radius_m)
  movel([0.229998, -1.347740, -2.593182, -0.771468, 1.570796, 1.800795],accel_mss,speed_ms,0,blend_radius_m)
  movel([0.230489, -1.348595, -2.592617, -0.771177, 1.570796, 1.801286],accel_mss,speed_ms,0,blend_radius_m)
  movel([0.230770, -1.349692, -2.591891, -0.770806, 1.570796, 1.801566],accel_mss,speed_ms,0,blend_radius_m)
  movel([0.230845, -1.350965, -2.591047, -0.770378, 1.570796, 1.801641],accel_mss,speed_ms,0,blend_radius_m)
  movel([0.230384, -1.354031, -2.589004, -0.769355, 1.570796, 1.801180],accel_mss,speed_ms,0,blend_radius_m)
  movel([0.229759, -1.356065, -2.587640, -0.768683, 1.570796, 1.800555],accel_mss,speed_ms,0,blend_radius_m)
  movel([0.228936, -1.358023, -2.586323, -0.768042, 1.570796, 1.799732],accel_mss,speed_ms,0,blend_radius_m)
  movel([0.227921, -1.359907, -2.585051, -0.767431, 1.570796, 1.798717],accel_mss,speed_ms,0,blend_radius_m)
  movel([0.226707, -1.361716, -2.583824, -0.766848, 1.570796, 1.797503],accel_mss,speed_ms,0,blend_radius_m)
  movel([0.225293, -1.363316, -2.582736, -0.766337, 1.570796, 1.796090],accel_mss,speed_ms,0,blend_radius_m)
  movel([0.223672, -1.364567, -2.581882, -0.765940, 1.570796, 1.794469],accel_mss,speed_ms,0,blend_radius_m)
  movel([0.221842, -1.365473, -2.581263, -0.765653, 1.570796, 1.792638],accel_mss,speed_ms,0,blend_radius_m)
  movel([0.219799, -1.366040, -2.580874, -0.765475, 1.570796, 1.790595],accel_mss,speed_ms,0,blend_radius_m)
  movel([0.218008, -1.366200, -2.580765, -0.765424, 1.570796, 1.788805],accel_mss,speed_ms,0,blend_radius_m)
  movel([0.216433, -1.365980, -2.580915, -0.765494, 1.570796, 1.787230],accel_mss,speed_ms,0,blend_radius_m)
  movel([0.215058, -1.365470, -2.581265, -0.765654, 1.570796, 1.785854],accel_mss,speed_ms,0,blend_radius_m)
  movel([0.213872, -1.364766, -2.581746, -0.765877, 1.570796, 1.784668],accel_mss,speed_ms,0,blend_radius_m)
  movel([0.211373, -1.362576, -2.583240, -0.766573, 1.570796, 1.782170],accel_mss,speed_ms,0,blend_radius_m)
  movel([0.208986, -1.360527, -2.584631, -0.767231, 1.570796, 1.779782],accel_mss,speed_ms,0,blend_radius_m)
  movel([0.207897, -1.359882, -2.585068, -0.767439, 1.570796, 1.778694],accel_mss,speed_ms,0,blend_radius_m)
  movel([0.206656, -1.359423, -2.585379, -0.767588, 1.570796, 1.777453],accel_mss,speed_ms,0,blend_radius_m)
  movel([0.205253, -1.359231, -2.585508, -0.767650, 1.570796, 1.776050],accel_mss,speed_ms,0,blend_radius_m)
  movel([0.203696, -1.359387, -2.585403, -0.767599, 1.570796, 1.774493],accel_mss,speed_ms,0,blend_radius_m)
  movel([0.203522, -1.360154, -2.584884, -0.767351, 1.570796, 1.774319],accel_mss,speed_ms,0,blend_radius_m)
  movel([0.203158, -1.362250, -2.583462, -0.766677, 1.570796, 1.773954],accel_mss,speed_ms,0,blend_radius_m)
  movel([0.203082, -1.364035, -2.582245, -0.766108, 1.570796, 1.773878],accel_mss,speed_ms,0,blend_radius_m)
  movel([0.203295, -1.365514, -2.581235, -0.765641, 1.570796, 1.774091],accel_mss,speed_ms,0,blend_radius_m)
  movel([0.203794, -1.366685, -2.580432, -0.765272, 1.570796, 1.774590],accel_mss,speed_ms,0,blend_radius_m)
  movel([0.204537, -1.367572, -2.579822, -0.764994, 1.570796, 1.775333],accel_mss,speed_ms,0,blend_radius_m)
  movel([0.205476, -1.368200, -2.579390, -0.764798, 1.570796, 1.776272],accel_mss,speed_ms,0,blend_radius_m)
  movel([0.206616, -1.368571, -2.579135, -0.764683, 1.570796, 1.777412],accel_mss,speed_ms,0,blend_radius_m)
  movel([0.207955, -1.368681, -2.579059, -0.764649, 1.570796, 1.778751],accel_mss,speed_ms,0,blend_radius_m)
  movel([0.200563, -1.370133, -2.578057, -0.764199, 1.570796, 1.771359],accel_mss,speed_ms,0,blend_radius_m)
  movel([0.205188, -1.349671, -2.591905, -0.770813, 1.570796, 1.775985],accel_mss,speed_ms,0,blend_radius_m)
  movel([0.205944, -1.349516, -2.592008, -0.770866, 1.570796, 1.776740],accel_mss,speed_ms,0,blend_radius_m)
  speed_ms = 0.003
  movel([0.205944, -1.342817, -2.588898, -0.780673, 1.570796, 1.776740],accel_mss,speed_ms,0,blend_radius_m)
  speed_ms = 1.000
  movel([0.205944, -1.317083, -2.576173, -0.819133, 1.570796, 1.776740],accel_mss,speed_ms,0,blend_radius_m)
  #M_RunCode9
  movel([0.204607, -1.339809, -2.561482, -0.811098, 1.570796, 1.775403],accel_mss,speed_ms,0,blend_radius_m)
  #M_RunCode3
  movel([0.204607, -1.365148, -2.573913, -0.773327, 1.570796, 1.775403],accel_mss,speed_ms,0,blend_radius_m)
  speed_ms = 0.003
  movel([0.204607, -1.371734, -2.576949, -0.763706, 1.570796, 1.775403],accel_mss,speed_ms,0,blend_radius_m)
  speed_ms = 0.007
  movel([0.205865, -1.371715, -2.576962, -0.763712, 1.570796, 1.776662],accel_mss,speed_ms,0,blend_radius_m)
  movel([0.206694, -1.372227, -2.576607, -0.763555, 1.570796, 1.777491],accel_mss,speed_ms,0,blend_radius_m)
  movel([0.207077, -1.373137, -2.575974, -0.763277, 1.570796, 1.777873],accel_mss,speed_ms,0,blend_radius_m)
  movel([0.207004, -1.374302, -2.575164, -0.762924, 1.570796, 1.777800],accel_mss,speed_ms,0,blend_radius_m)
  movel([0.206521, -1.375542, -2.574298, -0.762549, 1.570796, 1.777317],accel_mss,speed_ms,0,blend_radius_m)
  movel([0.205667, -1.376683, -2.573500, -0.762206, 1.570796, 1.776463],accel_mss,speed_ms,0,blend_radius_m)
  movel([0.204521, -1.377572, -2.572877, -0.761940, 1.570796, 1.775317],accel_mss,speed_ms,0,blend_radius_m)
  movel([0.203164, -1.378056, -2.572537, -0.761796, 1.570796, 1.773961],accel_mss,speed_ms,0,blend_radius_m)
  movel([0.202099, -1.378123, -2.572490, -0.761776, 1.570796, 1.772895],accel_mss,speed_ms,0,blend_radius_m)
  movel([0.201366, -1.377890, -2.572653, -0.761846, 1.570796, 1.772162],accel_mss,speed_ms,0,blend_radius_m)
  movel([0.200568, -1.377730, -2.572766, -0.761893, 1.570796, 1.771365],accel_mss,speed_ms,0,blend_radius_m)
  movel([0.199948, -1.377990, -2.572583, -0.761816, 1.570796, 1.770744],accel_mss,speed_ms,0,blend_radius_m)
  movel([0.199364, -1.378520, -2.572210, -0.761658, 1.570796, 1.770160],accel_mss,speed_ms,0,blend_radius_m)
  movel([0.198898, -1.379213, -2.571723, -0.761453, 1.570796, 1.769694],accel_mss,speed_ms,0,blend_radius_m)
  movel([0.198626, -1.379966, -2.571192, -0.761230, 1.570796, 1.769422],accel_mss,speed_ms,0,blend_radius_m)
  movel([0.198519, -1.380912, -2.570525, -0.760952, 1.570796, 1.769315],accel_mss,speed_ms,0,blend_radius_m)
  movel([0.198652, -1.381729, -2.569947, -0.760713, 1.570796, 1.769448],accel_mss,speed_ms,0,blend_radius_m)
  movel([0.199023, -1.382416, -2.569460, -0.760513, 1.570796, 1.769819],accel_mss,speed_ms,0,blend_radius_m)
  movel([0.199630, -1.382978, -2.569062, -0.760349, 1.570796, 1.770426],accel_mss,speed_ms,0,blend_radius_m)
  movel([0.200439, -1.383379, -2.568777, -0.760233, 1.570796, 1.771235],accel_mss,speed_ms,0,blend_radius_m)
  movel([0.201412, -1.383590, -2.568628, -0.760172, 1.570796, 1.772208],accel_mss,speed_ms,0,blend_radius_m)
  movel([0.202550, -1.383611, -2.568613, -0.760165, 1.570796, 1.773346],accel_mss,speed_ms,0,blend_radius_m)
  movel([0.203852, -1.383443, -2.568732, -0.760214, 1.570796, 1.774648],accel_mss,speed_ms,0,blend_radius_m)
  movel([0.206125, -1.382729, -2.569238, -0.760421, 1.570796, 1.776921],accel_mss,speed_ms,0,blend_radius_m)
  movel([0.208310, -1.381462, -2.570136, -0.760791, 1.570796, 1.779107],accel_mss,speed_ms,0,blend_radius_m)
  movel([0.209356, -1.380618, -2.570732, -0.761039, 1.570796, 1.780152],accel_mss,speed_ms,0,blend_radius_m)
  movel([0.210341, -1.379637, -2.571424, -0.761328, 1.570796, 1.781137],accel_mss,speed_ms,0,blend_radius_m)
  movel([0.212137, -1.377247, -2.573105, -0.762038, 1.570796, 1.782933],accel_mss,speed_ms,0,blend_radius_m)
  movel([0.213618, -1.374332, -2.575143, -0.762914, 1.570796, 1.784415],accel_mss,speed_ms,0,blend_radius_m)
  movel([0.214694, -1.370929, -2.577507, -0.763953, 1.570796, 1.785490],accel_mss,speed_ms,0,blend_radius_m)
  movel([0.225970, -1.368875, -2.578926, -0.764588, 1.570796, 1.796766],accel_mss,speed_ms,0,blend_radius_m)
  movel([0.222216, -1.383918, -2.568394, -0.760077, 1.570796, 1.793012],accel_mss,speed_ms,0,blend_radius_m)
  movel([0.214979, -1.385197, -2.567484, -0.759708, 1.570796, 1.785776],accel_mss,speed_ms,0,blend_radius_m)
  movel([0.216844, -1.384322, -2.568107, -0.759960, 1.570796, 1.787641],accel_mss,speed_ms,0,blend_radius_m)
  movel([0.218671, -1.383003, -2.569044, -0.760342, 1.570796, 1.789468],accel_mss,speed_ms,0,blend_radius_m)
  movel([0.220369, -1.381301, -2.570250, -0.760838, 1.570796, 1.791166],accel_mss,speed_ms,0,blend_radius_m)
  movel([0.221846, -1.379279, -2.571676, -0.761433, 1.570796, 1.792642],accel_mss,speed_ms,0,blend_radius_m)
  movel([0.223030, -1.377004, -2.573275, -0.762110, 1.570796, 1.793827],accel_mss,speed_ms,0,blend_radius_m)
  movel([0.223849, -1.374547, -2.574993, -0.762849, 1.570796, 1.794645],accel_mss,speed_ms,0,blend_radius_m)
  movel([0.215573, -1.376038, -2.573951, -0.762400, 1.570796, 1.786370],accel_mss,speed_ms,0,blend_radius_m)
  movel([0.214631, -1.379048, -2.571839, -0.761502, 1.570796, 1.785427],accel_mss,speed_ms,0,blend_radius_m)
  movel([0.213271, -1.382005, -2.569752, -0.760632, 1.570796, 1.784067],accel_mss,speed_ms,0,blend_radius_m)
  movel([0.211513, -1.384721, -2.567823, -0.759845, 1.570796, 1.782310],accel_mss,speed_ms,0,blend_radius_m)
  movel([0.210491, -1.385922, -2.566967, -0.759500, 1.570796, 1.781287],accel_mss,speed_ms,0,blend_radius_m)
  movel([0.209376, -1.387018, -2.566184, -0.759187, 1.570796, 1.780172],accel_mss,speed_ms,0,blend_radius_m)
  movel([0.208174, -1.387966, -2.565505, -0.758918, 1.570796, 1.778971],accel_mss,speed_ms,0,blend_radius_m)
  movel([0.206899, -1.388720, -2.564964, -0.758705, 1.570796, 1.777695],accel_mss,speed_ms,0,blend_radius_m)
  movel([0.205546, -1.389282, -2.564560, -0.758546, 1.570796, 1.776342],accel_mss,speed_ms,0,blend_radius_m)
  movel([0.204119, -1.389651, -2.564295, -0.758443, 1.570796, 1.774915],accel_mss,speed_ms,0,blend_radius_m)
  movel([0.202738, -1.389813, -2.564179, -0.758397, 1.570796, 1.773535],accel_mss,speed_ms,0,blend_radius_m)
  movel([0.201521, -1.389755, -2.564221, -0.758414, 1.570796, 1.772318],accel_mss,speed_ms,0,blend_radius_m)
  movel([0.200471, -1.389473, -2.564423, -0.758493, 1.570796, 1.771268],accel_mss,speed_ms,0,blend_radius_m)
  movel([0.199586, -1.388970, -2.564785, -0.758634, 1.570796, 1.770383],accel_mss,speed_ms,0,blend_radius_m)
  movel([0.198289, -1.387474, -2.565858, -0.759058, 1.570796, 1.769085],accel_mss,speed_ms,0,blend_radius_m)
  movel([0.197600, -1.385449, -2.567304, -0.759636, 1.570796, 1.768397],accel_mss,speed_ms,0,blend_radius_m)
  movel([0.197460, -1.383071, -2.568996, -0.760322, 1.570796, 1.768256],accel_mss,speed_ms,0,blend_radius_m)
  movel([0.197802, -1.380524, -2.570799, -0.761066, 1.570796, 1.768598],accel_mss,speed_ms,0,blend_radius_m)
  movel([0.198347, -1.378710, -2.572077, -0.761602, 1.570796, 1.769143],accel_mss,speed_ms,0,blend_radius_m)
  movel([0.199198, -1.376811, -2.573410, -0.762168, 1.570796, 1.769994],accel_mss,speed_ms,0,blend_radius_m)
  movel([0.200304, -1.375001, -2.574676, -0.762712, 1.570796, 1.771100],accel_mss,speed_ms,0,blend_radius_m)
  movel([0.201619, -1.373457, -2.575752, -0.763180, 1.570796, 1.772415],accel_mss,speed_ms,0,blend_radius_m)
  movel([0.203075, -1.372317, -2.576544, -0.763527, 1.570796, 1.773872],accel_mss,speed_ms,0,blend_radius_m)
  movel([0.204607, -1.371734, -2.576949, -0.763706, 1.570796, 1.775403],accel_mss,speed_ms,0,blend_radius_m)
  speed_ms = 0.003
  movel([0.204607, -1.365148, -2.573913, -0.773327, 1.570796, 1.775403],accel_mss,speed_ms,0,blend_radius_m)
  speed_ms = 1.000
  movel([0.204607, -1.339809, -2.561482, -0.811098, 1.570796, 1.775403],accel_mss,speed_ms,0,blend_radius_m)
  #M_RunCode9
  movel([0.281435, -1.240169, -2.621054, -0.851165, 1.570796, 1.852231],accel_mss,speed_ms,0,blend_radius_m)
  #M_RunCode3
  movel([0.281435, -1.267049, -2.634789, -0.810551, 1.570796, 1.852231],accel_mss,speed_ms,0,blend_radius_m)
  speed_ms = 0.003
  movel([0.281435, -1.274084, -2.638154, -0.800151, 1.570796, 1.852231],accel_mss,speed_ms,0,blend_radius_m)
  speed_ms = 0.007
  movel([0.281521, -1.274005, -2.638199, -0.800185, 1.570796, 1.852317],accel_mss,speed_ms,0,blend_radius_m)
  movel([0.281435, -1.274084, -2.638154, -0.800151, 1.570796, 1.852231],accel_mss,speed_ms,0,blend_radius_m)
  speed_ms = 0.003
  movel([0.281435, -1.267049, -2.634789, -0.810551, 1.570796, 1.852231],accel_mss,speed_ms,0,blend_radius_m)
  speed_ms = 1.000
  movel([0.281435, -1.240169, -2.621054, -0.851165, 1.570796, 1.852231],accel_mss,speed_ms,0,blend_radius_m)
  #M_RunCode9
  movel([0.257972, -1.256546, -2.612100, -0.843743, 1.570796, 1.828768],accel_mss,speed_ms,0,blend_radius_m)
  #M_RunCode3
  movel([0.257972, -1.283210, -2.625619, -0.803560, 1.570796, 1.828768],accel_mss,speed_ms,0,blend_radius_m)
  speed_ms = 0.003
  movel([0.257972, -1.290180, -2.628929, -0.793280, 1.570796, 1.828768],accel_mss,speed_ms,0,blend_radius_m)
  speed_ms = 0.007
  movel([0.258265, -1.291328, -2.628259, -0.792803, 1.570796, 1.829061],accel_mss,speed_ms,0,blend_radius_m)
  movel([0.258228, -1.292795, -2.627399, -0.792195, 1.570796, 1.829024],accel_mss,speed_ms,0,blend_radius_m)
  movel([0.257555, -1.295122, -2.626031, -0.791237, 1.570796, 1.828351],accel_mss,speed_ms,0,blend_radius_m)
  movel([0.256239, -1.297298, -2.624744, -0.790346, 1.570796, 1.827036],accel_mss,speed_ms,0,blend_radius_m)
  movel([0.254385, -1.299283, -2.623566, -0.789540, 1.570796, 1.825181],accel_mss,speed_ms,0,blend_radius_m)
  movel([0.252100, -1.301032, -2.622523, -0.788834, 1.570796, 1.822897],accel_mss,speed_ms,0,blend_radius_m)
  movel([0.249363, -1.302507, -2.621641, -0.788241, 1.570796, 1.820159],accel_mss,speed_ms,0,blend_radius_m)
  movel([0.246989, -1.303173, -2.621241, -0.787974, 1.570796, 1.817786],accel_mss,speed_ms,0,blend_radius_m)
  movel([0.244961, -1.303143, -2.621260, -0.787986, 1.570796, 1.815758],accel_mss,speed_ms,0,blend_radius_m)
  movel([0.243262, -1.302522, -2.621632, -0.788235, 1.570796, 1.814059],accel_mss,speed_ms,0,blend_radius_m)
  movel([0.241873, -1.301421, -2.622291, -0.788677, 1.570796, 1.812670],accel_mss,speed_ms,0,blend_radius_m)
  movel([0.240784, -1.299947, -2.623171, -0.789271, 1.570796, 1.811580],accel_mss,speed_ms,0,blend_radius_m)
  movel([0.239981, -1.298206, -2.624206, -0.789977, 1.570796, 1.810777],accel_mss,speed_ms,0,blend_radius_m)
  movel([0.239453, -1.296304, -2.625333, -0.790752, 1.570796, 1.810249],accel_mss,speed_ms,0,blend_radius_m)
  movel([0.241828, -1.294022, -2.626678, -0.791689, 1.570796, 1.812625],accel_mss,speed_ms,0,blend_radius_m)
  movel([0.244783, -1.291914, -2.627916, -0.792559, 1.570796, 1.815579],accel_mss,speed_ms,0,blend_radius_m)
  movel([0.248026, -1.290158, -2.628942, -0.793289, 1.570796, 1.818822],accel_mss,speed_ms,0,blend_radius_m)
  movel([0.251261, -1.288932, -2.629656, -0.793801, 1.570796, 1.822057],accel_mss,speed_ms,0,blend_radius_m)
  movel([0.254197, -1.288411, -2.629959, -0.794019, 1.570796, 1.824993],accel_mss,speed_ms,0,blend_radius_m)
  movel([0.255457, -1.288472, -2.629923, -0.793993, 1.570796, 1.826254],accel_mss,speed_ms,0,blend_radius_m)
  movel([0.256532, -1.288772, -2.629749, -0.793868, 1.570796, 1.827328],accel_mss,speed_ms,0,blend_radius_m)
  movel([0.257381, -1.289335, -2.629422, -0.793633, 1.570796, 1.828178],accel_mss,speed_ms,0,blend_radius_m)
  movel([0.257972, -1.290180, -2.628929, -0.793280, 1.570796, 1.828768],accel_mss,speed_ms,0,blend_radius_m)
  speed_ms = 0.003
  movel([0.257972, -1.283210, -2.625619, -0.803560, 1.570796, 1.828768],accel_mss,speed_ms,0,blend_radius_m)
  speed_ms = 1.000
  movel([0.257972, -1.256546, -2.612100, -0.843743, 1.570796, 1.828768],accel_mss,speed_ms,0,blend_radius_m)
  #M_RunCode9
  movel([0.324800, -1.226006, -2.628547, -0.857837, 1.570796, 1.895597],accel_mss,speed_ms,0,blend_radius_m)
  #M_RunCode3
  movel([0.324800, -1.253058, -2.642469, -0.816862, 1.570796, 1.895597],accel_mss,speed_ms,0,blend_radius_m)
  speed_ms = 0.003
  movel([0.324800, -1.260146, -2.645882, -0.806361, 1.570796, 1.895597],accel_mss,speed_ms,0,blend_radius_m)
  speed_ms = 0.007
  movel([0.325189, -1.258580, -2.646735, -0.807073, 1.570796, 1.895986],accel_mss,speed_ms,0,blend_radius_m)
  movel([0.325795, -1.256940, -2.647626, -0.807823, 1.570796, 1.896591],accel_mss,speed_ms,0,blend_radius_m)
  movel([0.326278, -1.257078, -2.647551, -0.807760, 1.570796, 1.897074],accel_mss,speed_ms,0,blend_radius_m)
  movel([0.326346, -1.257559, -2.647290, -0.807540, 1.570796, 1.897142],accel_mss,speed_ms,0,blend_radius_m)
  movel([0.326468, -1.258090, -2.647002, -0.807297, 1.570796, 1.897264],accel_mss,speed_ms,0,blend_radius_m)
  movel([0.327111, -1.258378, -2.646845, -0.807165, 1.570796, 1.897908],accel_mss,speed_ms,0,blend_radius_m)
  movel([0.328054, -1.258279, -2.646899, -0.807211, 1.570796, 1.898850],accel_mss,speed_ms,0,blend_radius_m)
  movel([0.329072, -1.257962, -2.647072, -0.807356, 1.570796, 1.899869],accel_mss,speed_ms,0,blend_radius_m)
  movel([0.330498, -1.257467, -2.647340, -0.807582, 1.570796, 1.901294],accel_mss,speed_ms,0,blend_radius_m)
  movel([0.331361, -1.255398, -2.648460, -0.808531, 1.570796, 1.902157],accel_mss,speed_ms,0,blend_radius_m)
  movel([0.331584, -1.253748, -2.649350, -0.809291, 1.570796, 1.902380],accel_mss,speed_ms,0,blend_radius_m)
  movel([0.331375, -1.253153, -2.649670, -0.809566, 1.570796, 1.902171],accel_mss,speed_ms,0,blend_radius_m)
  movel([0.330915, -1.252750, -2.649887, -0.809753, 1.570796, 1.901712],accel_mss,speed_ms,0,blend_radius_m)
  movel([0.330170, -1.252567, -2.649985, -0.809837, 1.570796, 1.900966],accel_mss,speed_ms,0,blend_radius_m)
  movel([0.329109, -1.252637, -2.649947, -0.809805, 1.570796, 1.899905],accel_mss,speed_ms,0,blend_radius_m)
  movel([0.330088, -1.251538, -2.650536, -0.810315, 1.570796, 1.900885],accel_mss,speed_ms,0,blend_radius_m)
  movel([0.331013, -1.250665, -2.651003, -0.810720, 1.570796, 1.901810],accel_mss,speed_ms,0,blend_radius_m)
  movel([0.331423, -1.250432, -2.651128, -0.810829, 1.570796, 1.902219],accel_mss,speed_ms,0,blend_radius_m)
  movel([0.331777, -1.250392, -2.651149, -0.810848, 1.570796, 1.902573],accel_mss,speed_ms,0,blend_radius_m)
  movel([0.332271, -1.251081, -2.650781, -0.810527, 1.570796, 1.903067],accel_mss,speed_ms,0,blend_radius_m)
  movel([0.332492, -1.253102, -2.649697, -0.809590, 1.570796, 1.903288],accel_mss,speed_ms,0,blend_radius_m)
  movel([0.332162, -1.255402, -2.648458, -0.808529, 1.570796, 1.902959],accel_mss,speed_ms,0,blend_radius_m)
  movel([0.331744, -1.256560, -2.647832, -0.807997, 1.570796, 1.902541],accel_mss,speed_ms,0,blend_radius_m)
  movel([0.331127, -1.257674, -2.647228, -0.807487, 1.570796, 1.901923],accel_mss,speed_ms,0,blend_radius_m)
  movel([0.330293, -1.258704, -2.646668, -0.807017, 1.570796, 1.901089],accel_mss,speed_ms,0,blend_radius_m)
  movel([0.329221, -1.259614, -2.646172, -0.806603, 1.570796, 1.900017],accel_mss,speed_ms,0,blend_radius_m)
  movel([0.329024, -1.258380, -2.646844, -0.807164, 1.570796, 1.899820],accel_mss,speed_ms,0,blend_radius_m)
  movel([0.325403, -1.262656, -2.644508, -0.805225, 1.570796, 1.896199],accel_mss,speed_ms,0,blend_radius_m)
  movel([0.324812, -1.261539, -2.645121, -0.805730, 1.570796, 1.895608],accel_mss,speed_ms,0,blend_radius_m)
  movel([0.324800, -1.260146, -2.645882, -0.806361, 1.570796, 1.895597],accel_mss,speed_ms,0,blend_radius_m)
  speed_ms = 0.003
  movel([0.324800, -1.253058, -2.642469, -0.816862, 1.570796, 1.895597],accel_mss,speed_ms,0,blend_radius_m)
  speed_ms = 1.000
  movel([0.324800, -1.226006, -2.628547, -0.857837, 1.570796, 1.895597],accel_mss,speed_ms,0,blend_radius_m)
  #M_RunCode9
  movel([0.334430, -1.184074, -2.649412, -0.878903, 1.570796, 1.905226],accel_mss,speed_ms,0,blend_radius_m)
  #M_RunCode3
  movel([0.334430, -1.211558, -2.663890, -0.836941, 1.570796, 1.905226],accel_mss,speed_ms,0,blend_radius_m)
  speed_ms = 0.003
  movel([0.334430, -1.218783, -2.667445, -0.826162, 1.570796, 1.905226],accel_mss,speed_ms,0,blend_radius_m)
  speed_ms = 0.007
  movel([0.332348, -1.219318, -2.667178, -0.825892, 1.570796, 1.903144],accel_mss,speed_ms,0,blend_radius_m)
  movel([0.330315, -1.219605, -2.667035, -0.825749, 1.570796, 1.901112],accel_mss,speed_ms,0,blend_radius_m)
  movel([0.328361, -1.219627, -2.667024, -0.825737, 1.570796, 1.899157],accel_mss,speed_ms,0,blend_radius_m)
  movel([0.326513, -1.219367, -2.667154, -0.825868, 1.570796, 1.897309],accel_mss,speed_ms,0,blend_radius_m)
  movel([0.324802, -1.218813, -2.667429, -0.826146, 1.570796, 1.895598],accel_mss,speed_ms,0,blend_radius_m)
  movel([0.324085, -1.218270, -2.667699, -0.826420, 1.570796, 1.894881],accel_mss,speed_ms,0,blend_radius_m)
  movel([0.323480, -1.217525, -2.668069, -0.826795, 1.570796, 1.894276],accel_mss,speed_ms,0,blend_radius_m)
  movel([0.322934, -1.216862, -2.668398, -0.827130, 1.570796, 1.893730],accel_mss,speed_ms,0,blend_radius_m)
  movel([0.322382, -1.216563, -2.668545, -0.827280, 1.570796, 1.893178],accel_mss,speed_ms,0,blend_radius_m)
  movel([0.321004, -1.216860, -2.668399, -0.827130, 1.570796, 1.891800],accel_mss,speed_ms,0,blend_radius_m)
  movel([0.319016, -1.217575, -2.668044, -0.826770, 1.570796, 1.889812],accel_mss,speed_ms,0,blend_radius_m)
  movel([0.316929, -1.218353, -2.667658, -0.826378, 1.570796, 1.887726],accel_mss,speed_ms,0,blend_radius_m)
  movel([0.315257, -1.218834, -2.667419, -0.826136, 1.570796, 1.886054],accel_mss,speed_ms,0,blend_radius_m)
  movel([0.312327, -1.219080, -2.667297, -0.826012, 1.570796, 1.883124],accel_mss,speed_ms,0,blend_radius_m)
  movel([0.309978, -1.218785, -2.667444, -0.826161, 1.570796, 1.880774],accel_mss,speed_ms,0,blend_radius_m)
  movel([0.308157, -1.218003, -2.667832, -0.826554, 1.570796, 1.878953],accel_mss,speed_ms,0,blend_radius_m)
  movel([0.306816, -1.216786, -2.668435, -0.827168, 1.570796, 1.877612],accel_mss,speed_ms,0,blend_radius_m)
  movel([0.305908, -1.215177, -2.669230, -0.827982, 1.570796, 1.876705],accel_mss,speed_ms,0,blend_radius_m)
  movel([0.305384, -1.213233, -2.670187, -0.828969, 1.570796, 1.876181],accel_mss,speed_ms,0,blend_radius_m)
  movel([0.305199, -1.211003, -2.671279, -0.830107, 1.570796, 1.875995],accel_mss,speed_ms,0,blend_radius_m)
  movel([0.305299, -1.208535, -2.672481, -0.831373, 1.570796, 1.876096],accel_mss,speed_ms,0,blend_radius_m)
  movel([0.306177, -1.203106, -2.675102, -0.834182, 1.570796, 1.876974],accel_mss,speed_ms,0,blend_radius_m)
  movel([0.307636, -1.197368, -2.677836, -0.837185, 1.570796, 1.878432],accel_mss,speed_ms,0,blend_radius_m)
  movel([0.310678, -1.186775, -2.682789, -0.842825, 1.570796, 1.881474],accel_mss,speed_ms,0,blend_radius_m)
  movel([0.311637, -1.182182, -2.684900, -0.845308, 1.570796, 1.882433],accel_mss,speed_ms,0,blend_radius_m)
  movel([0.312334, -1.176967, -2.687268, -0.848154, 1.570796, 1.883130],accel_mss,speed_ms,0,blend_radius_m)
  movel([0.312710, -1.171412, -2.689760, -0.851217, 1.570796, 1.883506],accel_mss,speed_ms,0,blend_radius_m)
  movel([0.312704, -1.165797, -2.692245, -0.854346, 1.570796, 1.883500],accel_mss,speed_ms,0,blend_radius_m)
  movel([0.312245, -1.160421, -2.694595, -0.857373, 1.570796, 1.883042],accel_mss,speed_ms,0,blend_radius_m)
  movel([0.311269, -1.155584, -2.696684, -0.860122, 1.570796, 1.882065],accel_mss,speed_ms,0,blend_radius_m)
  movel([0.309710, -1.151600, -2.698386, -0.862403, 1.570796, 1.880506],accel_mss,speed_ms,0,blend_radius_m)
  movel([0.308692, -1.150028, -2.699053, -0.863307, 1.570796, 1.879489],accel_mss,speed_ms,0,blend_radius_m)
  movel([0.307505, -1.148786, -2.699579, -0.864024, 1.570796, 1.878302],accel_mss,speed_ms,0,blend_radius_m)
  movel([0.306038, -1.147782, -2.700003, -0.864605, 1.570796, 1.876834],accel_mss,speed_ms,0,blend_radius_m)
  movel([0.304105, -1.146877, -2.700384, -0.865129, 1.570796, 1.874901],accel_mss,speed_ms,0,blend_radius_m)
  movel([0.301771, -1.146197, -2.700669, -0.865523, 1.570796, 1.872567],accel_mss,speed_ms,0,blend_radius_m)
  movel([0.299106, -1.145864, -2.700809, -0.865716, 1.570796, 1.869903],accel_mss,speed_ms,0,blend_radius_m)
  movel([0.296181, -1.146006, -2.700750, -0.865633, 1.570796, 1.866977],accel_mss,speed_ms,0,blend_radius_m)
  movel([0.293066, -1.146740, -2.700441, -0.865208, 1.570796, 1.863863],accel_mss,speed_ms,0,blend_radius_m)
  movel([0.289839, -1.148186, -2.699832, -0.864371, 1.570796, 1.860636],accel_mss,speed_ms,0,blend_radius_m)
  movel([0.288206, -1.149214, -2.699398, -0.863777, 1.570796, 1.859003],accel_mss,speed_ms,0,blend_radius_m)
  movel([0.286575, -1.150459, -2.698871, -0.863059, 1.570796, 1.857371],accel_mss,speed_ms,0,blend_radius_m)
  movel([0.284270, -1.152720, -2.697909, -0.861760, 1.570796, 1.855066],accel_mss,speed_ms,0,blend_radius_m)
  movel([0.282632, -1.155047, -2.696914, -0.860428, 1.570796, 1.853428],accel_mss,speed_ms,0,blend_radius_m)
  movel([0.281596, -1.157415, -2.695896, -0.859078, 1.570796, 1.852392],accel_mss,speed_ms,0,blend_radius_m)
  movel([0.281094, -1.159808, -2.694861, -0.857720, 1.570796, 1.851891],accel_mss,speed_ms,0,blend_radius_m)
  movel([0.281065, -1.162206, -2.693818, -0.856365, 1.570796, 1.851861],accel_mss,speed_ms,0,blend_radius_m)
  movel([0.281434, -1.164600, -2.692771, -0.855018, 1.570796, 1.852231],accel_mss,speed_ms,0,blend_radius_m)
  movel([0.282136, -1.166969, -2.691729, -0.853690, 1.570796, 1.852933],accel_mss,speed_ms,0,blend_radius_m)
  movel([0.283109, -1.169300, -2.690698, -0.852390, 1.570796, 1.853905],accel_mss,speed_ms,0,blend_radius_m)
  movel([0.285594, -1.173786, -2.688699, -0.849904, 1.570796, 1.856391],accel_mss,speed_ms,0,blend_radius_m)
  movel([0.288387, -1.177926, -2.686835, -0.847628, 1.570796, 1.859183],accel_mss,speed_ms,0,blend_radius_m)
  movel([0.290989, -1.181581, -2.685174, -0.845634, 1.570796, 1.861785],accel_mss,speed_ms,0,blend_radius_m)
  movel([0.292912, -1.184613, -2.683785, -0.843990, 1.570796, 1.863708],accel_mss,speed_ms,0,blend_radius_m)
  movel([0.297110, -1.192274, -2.680233, -0.839882, 1.570796, 1.867906],accel_mss,speed_ms,0,blend_radius_m)
  movel([0.299195, -1.196465, -2.678263, -0.837661, 1.570796, 1.869991],accel_mss,speed_ms,0,blend_radius_m)
  movel([0.300532, -1.199948, -2.676611, -0.835830, 1.570796, 1.871328],accel_mss,speed_ms,0,blend_radius_m)
  movel([0.300808, -1.201478, -2.675881, -0.835030, 1.570796, 1.871604],accel_mss,speed_ms,0,blend_radius_m)
  movel([0.300849, -1.203096, -2.675107, -0.834187, 1.570796, 1.871646],accel_mss,speed_ms,0,blend_radius_m)
  movel([0.300291, -1.206550, -2.673443, -0.832396, 1.570796, 1.871087],accel_mss,speed_ms,0,blend_radius_m)
  movel([0.298982, -1.210187, -2.671677, -0.830525, 1.570796, 1.869779],accel_mss,speed_ms,0,blend_radius_m)
  movel([0.297057, -1.213892, -2.669863, -0.828634, 1.570796, 1.867854],accel_mss,speed_ms,0,blend_radius_m)
  movel([0.294638, -1.217549, -2.668057, -0.826783, 1.570796, 1.865435],accel_mss,speed_ms,0,blend_radius_m)
  movel([0.291848, -1.221051, -2.666314, -0.825024, 1.570796, 1.862644],accel_mss,speed_ms,0,blend_radius_m)
  movel([0.288802, -1.224288, -2.664690, -0.823411, 1.570796, 1.859599],accel_mss,speed_ms,0,blend_radius_m)
  movel([0.285623, -1.227158, -2.663240, -0.821991, 1.570796, 1.856419],accel_mss,speed_ms,0,blend_radius_m)
  movel([0.281531, -1.230193, -2.661696, -0.820499, 1.570796, 1.852328],accel_mss,speed_ms,0,blend_radius_m)
  movel([0.279753, -1.231241, -2.661161, -0.819987, 1.570796, 1.850550],accel_mss,speed_ms,0,blend_radius_m)
  movel([0.278125, -1.232014, -2.660765, -0.819610, 1.570796, 1.848921],accel_mss,speed_ms,0,blend_radius_m)
  movel([0.276626, -1.232539, -2.660496, -0.819354, 1.570796, 1.847423],accel_mss,speed_ms,0,blend_radius_m)
  movel([0.275229, -1.232844, -2.660339, -0.819205, 1.570796, 1.846026],accel_mss,speed_ms,0,blend_radius_m)
  movel([0.272671, -1.232889, -2.660316, -0.819184, 1.570796, 1.843467],accel_mss,speed_ms,0,blend_radius_m)
  movel([0.270277, -1.232363, -2.660587, -0.819440, 1.570796, 1.841073],accel_mss,speed_ms,0,blend_radius_m)
  movel([0.267886, -1.231472, -2.661043, -0.819874, 1.570796, 1.838682],accel_mss,speed_ms,0,blend_radius_m)
  movel([0.262441, -1.229432, -2.662084, -0.820872, 1.570796, 1.833238],accel_mss,speed_ms,0,blend_radius_m)
  movel([0.262136, -1.229362, -2.662120, -0.820907, 1.570796, 1.832932],accel_mss,speed_ms,0,blend_radius_m)
  movel([0.262160, -1.229515, -2.662042, -0.820832, 1.570796, 1.832956],accel_mss,speed_ms,0,blend_radius_m)
  movel([0.263010, -1.230374, -2.661604, -0.820411, 1.570796, 1.833806],accel_mss,speed_ms,0,blend_radius_m)
  movel([0.266750, -1.233473, -2.660016, -0.818900, 1.570796, 1.837547],accel_mss,speed_ms,0,blend_radius_m)
  movel([0.272915, -1.238617, -2.657356, -0.816416, 1.570796, 1.843712],accel_mss,speed_ms,0,blend_radius_m)
  movel([0.267662, -1.238476, -2.657429, -0.816483, 1.570796, 1.838458],accel_mss,speed_ms,0,blend_radius_m)
  movel([0.261977, -1.237989, -2.657682, -0.816717, 1.570796, 1.832773],accel_mss,speed_ms,0,blend_radius_m)
  movel([0.256038, -1.237218, -2.658083, -0.817088, 1.570796, 1.826835],accel_mss,speed_ms,0,blend_radius_m)
  movel([0.250020, -1.236226, -2.658597, -0.817567, 1.570796, 1.820817],accel_mss,speed_ms,0,blend_radius_m)
  movel([0.238492, -1.233772, -2.659862, -0.818754, 1.570796, 1.809288],accel_mss,speed_ms,0,blend_radius_m)
  movel([0.233360, -1.232403, -2.660566, -0.819420, 1.570796, 1.804156],accel_mss,speed_ms,0,blend_radius_m)
  movel([0.228912, -1.230987, -2.661291, -0.820111, 1.570796, 1.799708],accel_mss,speed_ms,0,blend_radius_m)
  movel([0.220613, -1.232516, -2.660508, -0.819365, 1.570796, 1.791409],accel_mss,speed_ms,0,blend_radius_m)
  movel([0.211878, -1.234584, -2.659444, -0.818360, 1.570796, 1.782675],accel_mss,speed_ms,0,blend_radius_m)
  movel([0.193790, -1.239544, -2.656873, -0.815972, 1.570796, 1.764586],accel_mss,speed_ms,0,blend_radius_m)
  movel([0.184758, -1.242046, -2.655566, -0.814777, 1.570796, 1.755554],accel_mss,speed_ms,0,blend_radius_m)
  movel([0.175945, -1.244302, -2.654380, -0.813707, 1.570796, 1.746741],accel_mss,speed_ms,0,blend_radius_m)
  movel([0.167493, -1.246114, -2.653423, -0.812852, 1.570796, 1.738290],accel_mss,speed_ms,0,blend_radius_m)
  movel([0.159544, -1.247293, -2.652799, -0.812297, 1.570796, 1.730340],accel_mss,speed_ms,0,blend_radius_m)
  movel([0.156613, -1.247470, -2.652705, -0.812214, 1.570796, 1.727409],accel_mss,speed_ms,0,blend_radius_m)
  movel([0.153986, -1.247367, -2.652759, -0.812262, 1.570796, 1.724783],accel_mss,speed_ms,0,blend_radius_m)
  movel([0.151672, -1.246994, -2.652958, -0.812438, 1.570796, 1.722469],accel_mss,speed_ms,0,blend_radius_m)
  movel([0.149679, -1.246362, -2.653292, -0.812735, 1.570796, 1.720475],accel_mss,speed_ms,0,blend_radius_m)
  movel([0.148018, -1.245478, -2.653759, -0.813151, 1.570796, 1.718814],accel_mss,speed_ms,0,blend_radius_m)
  movel([0.146696, -1.244357, -2.654351, -0.813681, 1.570796, 1.717492],accel_mss,speed_ms,0,blend_radius_m)
  movel([0.145729, -1.243000, -2.655065, -0.814324, 1.570796, 1.716526],accel_mss,speed_ms,0,blend_radius_m)
  movel([0.145126, -1.241419, -2.655894, -0.815076, 1.570796, 1.715922],accel_mss,speed_ms,0,blend_radius_m)
  movel([0.144899, -1.239626, -2.656830, -0.815932, 1.570796, 1.715696],accel_mss,speed_ms,0,blend_radius_m)
  movel([0.145064, -1.237627, -2.657871, -0.816892, 1.570796, 1.715861],accel_mss,speed_ms,0,blend_radius_m)
  movel([0.145630, -1.235428, -2.659009, -0.817952, 1.570796, 1.716427],accel_mss,speed_ms,0,blend_radius_m)
  movel([0.146612, -1.233043, -2.660237, -0.819108, 1.570796, 1.717409],accel_mss,speed_ms,0,blend_radius_m)
  movel([0.148023, -1.230482, -2.661549, -0.820358, 1.570796, 1.718819],accel_mss,speed_ms,0,blend_radius_m)
  movel([0.149875, -1.227751, -2.662939, -0.821699, 1.570796, 1.720672],accel_mss,speed_ms,0,blend_radius_m)
  movel([0.152186, -1.224864, -2.664400, -0.823125, 1.570796, 1.722982],accel_mss,speed_ms,0,blend_radius_m)
  movel([0.154968, -1.221827, -2.665926, -0.824637, 1.570796, 1.725765],accel_mss,speed_ms,0,blend_radius_m)
  movel([0.155699, -1.224272, -2.664698, -0.823419, 1.570796, 1.726495],accel_mss,speed_ms,0,blend_radius_m)
  movel([0.156145, -1.225396, -2.664131, -0.822861, 1.570796, 1.726942],accel_mss,speed_ms,0,blend_radius_m)
  movel([0.156901, -1.226200, -2.663725, -0.822464, 1.570796, 1.727697],accel_mss,speed_ms,0,blend_radius_m)
  movel([0.157823, -1.226462, -2.663593, -0.822335, 1.570796, 1.728619],accel_mss,speed_ms,0,blend_radius_m)
  movel([0.159170, -1.226459, -2.663594, -0.822336, 1.570796, 1.729966],accel_mss,speed_ms,0,blend_radius_m)
  movel([0.162914, -1.225780, -2.663937, -0.822672, 1.570796, 1.733710],accel_mss,speed_ms,0,blend_radius_m)
  movel([0.167690, -1.224417, -2.664625, -0.823347, 1.570796, 1.738487],accel_mss,speed_ms,0,blend_radius_m)
  movel([0.173067, -1.222608, -2.665534, -0.824247, 1.570796, 1.743863],accel_mss,speed_ms,0,blend_radius_m)
  movel([0.183836, -1.218644, -2.667513, -0.826231, 1.570796, 1.754632],accel_mss,speed_ms,0,blend_radius_m)
  movel([0.191621, -1.215793, -2.668926, -0.827670, 1.570796, 1.762417],accel_mss,speed_ms,0,blend_radius_m)
  movel([0.198193, -1.213897, -2.669860, -0.828631, 1.570796, 1.768990],accel_mss,speed_ms,0,blend_radius_m)
  movel([0.204768, -1.212036, -2.670774, -0.829580, 1.570796, 1.775564],accel_mss,speed_ms,0,blend_radius_m)
  movel([0.196265, -1.207748, -2.672863, -0.831778, 1.570796, 1.767061],accel_mss,speed_ms,0,blend_radius_m)
  movel([0.192039, -1.205222, -2.674084, -0.833083, 1.570796, 1.762836],accel_mss,speed_ms,0,blend_radius_m)
  movel([0.188387, -1.202195, -2.675538, -0.834656, 1.570796, 1.759183],accel_mss,speed_ms,0,blend_radius_m)
  movel([0.186912, -1.200428, -2.676382, -0.835579, 1.570796, 1.757709],accel_mss,speed_ms,0,blend_radius_m)
  movel([0.185741, -1.198455, -2.677321, -0.836613, 1.570796, 1.756538],accel_mss,speed_ms,0,blend_radius_m)
  movel([0.184931, -1.196253, -2.678363, -0.837773, 1.570796, 1.755728],accel_mss,speed_ms,0,blend_radius_m)
  movel([0.184540, -1.193788, -2.679523, -0.839077, 1.570796, 1.755336],accel_mss,speed_ms,0,blend_radius_m)
  movel([0.184621, -1.191036, -2.680811, -0.840542, 1.570796, 1.755418],accel_mss,speed_ms,0,blend_radius_m)
  movel([0.185234, -1.187966, -2.682239, -0.842185, 1.570796, 1.756030],accel_mss,speed_ms,0,blend_radius_m)
  movel([0.186438, -1.184546, -2.683816, -0.844027, 1.570796, 1.757234],accel_mss,speed_ms,0,blend_radius_m)
  movel([0.188295, -1.180746, -2.685554, -0.846088, 1.570796, 1.759092],accel_mss,speed_ms,0,blend_radius_m)
  movel([0.191123, -1.176312, -2.687564, -0.848513, 1.570796, 1.761919],accel_mss,speed_ms,0,blend_radius_m)
  movel([0.194627, -1.171957, -2.689517, -0.850915, 1.570796, 1.765423],accel_mss,speed_ms,0,blend_radius_m)
  movel([0.198669, -1.167808, -2.691359, -0.853222, 1.570796, 1.769465],accel_mss,speed_ms,0,blend_radius_m)
  movel([0.203104, -1.163993, -2.693037, -0.855359, 1.570796, 1.773900],accel_mss,speed_ms,0,blend_radius_m)
  movel([0.207785, -1.160640, -2.694500, -0.857249, 1.570796, 1.778581],accel_mss,speed_ms,0,blend_radius_m)
  movel([0.212561, -1.157886, -2.695692, -0.858810, 1.570796, 1.783358],accel_mss,speed_ms,0,blend_radius_m)
  movel([0.217275, -1.155865, -2.696563, -0.859961, 1.570796, 1.788071],accel_mss,speed_ms,0,blend_radius_m)
  movel([0.221766, -1.154703, -2.697061, -0.860625, 1.570796, 1.792562],accel_mss,speed_ms,0,blend_radius_m)
  movel([0.223897, -1.154756, -2.697039, -0.860594, 1.570796, 1.794693],accel_mss,speed_ms,0,blend_radius_m)
  movel([0.225887, -1.155437, -2.696747, -0.860205, 1.570796, 1.796684],accel_mss,speed_ms,0,blend_radius_m)
  movel([0.227070, -1.156576, -2.696257, -0.859556, 1.570796, 1.797867],accel_mss,speed_ms,0,blend_radius_m)
  movel([0.227153, -1.157267, -2.695959, -0.859162, 1.570796, 1.797949],accel_mss,speed_ms,0,blend_radius_m)
  movel([0.226782, -1.158010, -2.695639, -0.858740, 1.570796, 1.797578],accel_mss,speed_ms,0,blend_radius_m)
  movel([0.225235, -1.157437, -2.695886, -0.859066, 1.570796, 1.796032],accel_mss,speed_ms,0,blend_radius_m)
  movel([0.223752, -1.157201, -2.695988, -0.859200, 1.570796, 1.794548],accel_mss,speed_ms,0,blend_radius_m)
  movel([0.222348, -1.157272, -2.695957, -0.859159, 1.570796, 1.793144],accel_mss,speed_ms,0,blend_radius_m)
  movel([0.221029, -1.157620, -2.695807, -0.858962, 1.570796, 1.791826],accel_mss,speed_ms,0,blend_radius_m)
  movel([0.219806, -1.158215, -2.695550, -0.858623, 1.570796, 1.790603],accel_mss,speed_ms,0,blend_radius_m)
  movel([0.218686, -1.159030, -2.695198, -0.858161, 1.570796, 1.789482],accel_mss,speed_ms,0,blend_radius_m)
  movel([0.217682, -1.160031, -2.694764, -0.857594, 1.570796, 1.788479],accel_mss,speed_ms,0,blend_radius_m)
  movel([0.216806, -1.161186, -2.694263, -0.856941, 1.570796, 1.787602],accel_mss,speed_ms,0,blend_radius_m)
  movel([0.215449, -1.163853, -2.693099, -0.855437, 1.570796, 1.786246],accel_mss,speed_ms,0,blend_radius_m)
  movel([0.214692, -1.166790, -2.691808, -0.853790, 1.570796, 1.785488],accel_mss,speed_ms,0,blend_radius_m)
  movel([0.214585, -1.169780, -2.690486, -0.852124, 1.570796, 1.785381],accel_mss,speed_ms,0,blend_radius_m)
  movel([0.215194, -1.172589, -2.689235, -0.850566, 1.570796, 1.785991],accel_mss,speed_ms,0,blend_radius_m)
  movel([0.215946, -1.174002, -2.688602, -0.849785, 1.570796, 1.786743],accel_mss,speed_ms,0,blend_radius_m)
  movel([0.217130, -1.175452, -2.687951, -0.848986, 1.570796, 1.787926],accel_mss,speed_ms,0,blend_radius_m)
  movel([0.220571, -1.178414, -2.686614, -0.847361, 1.570796, 1.791368],accel_mss,speed_ms,0,blend_radius_m)
  movel([0.225076, -1.181399, -2.685257, -0.845733, 1.570796, 1.795873],accel_mss,speed_ms,0,blend_radius_m)
  movel([0.230207, -1.184315, -2.683922, -0.844152, 1.570796, 1.801003],accel_mss,speed_ms,0,blend_radius_m)
  movel([0.240675, -1.189549, -2.681504, -0.841336, 1.570796, 1.811471],accel_mss,speed_ms,0,blend_radius_m)
  movel([0.248737, -1.193195, -2.679802, -0.839392, 1.570796, 1.819534],accel_mss,speed_ms,0,blend_radius_m)
  movel([0.252795, -1.195003, -2.678952, -0.838433, 1.570796, 1.823591],accel_mss,speed_ms,0,blend_radius_m)
  movel([0.255056, -1.195864, -2.678546, -0.837978, 1.570796, 1.825852],accel_mss,speed_ms,0,blend_radius_m)
  movel([0.256928, -1.196287, -2.678347, -0.837755, 1.570796, 1.827725],accel_mss,speed_ms,0,blend_radius_m)
  movel([0.257538, -1.196247, -2.678366, -0.837776, 1.570796, 1.828334],accel_mss,speed_ms,0,blend_radius_m)
  movel([0.257911, -1.196022, -2.678472, -0.837895, 1.570796, 1.828707],accel_mss,speed_ms,0,blend_radius_m)
  movel([0.258248, -1.194987, -2.678960, -0.838442, 1.570796, 1.829044],accel_mss,speed_ms,0,blend_radius_m)
  movel([0.258310, -1.192212, -2.680262, -0.839915, 1.570796, 1.829106],accel_mss,speed_ms,0,blend_radius_m)
  movel([0.257837, -1.189604, -2.681478, -0.841307, 1.570796, 1.828633],accel_mss,speed_ms,0,blend_radius_m)
  movel([0.256524, -1.184157, -2.683995, -0.844237, 1.570796, 1.827321],accel_mss,speed_ms,0,blend_radius_m)
  movel([0.256319, -1.180944, -2.685464, -0.845981, 1.570796, 1.827116],accel_mss,speed_ms,0,blend_radius_m)
  movel([0.256842, -1.177141, -2.687190, -0.848058, 1.570796, 1.827639],accel_mss,speed_ms,0,blend_radius_m)
  movel([0.257482, -1.174955, -2.688175, -0.849260, 1.570796, 1.828278],accel_mss,speed_ms,0,blend_radius_m)
  movel([0.258431, -1.172542, -2.689255, -0.850591, 1.570796, 1.829227],accel_mss,speed_ms,0,blend_radius_m)
  movel([0.259727, -1.169878, -2.690442, -0.852069, 1.570796, 1.830523],accel_mss,speed_ms,0,blend_radius_m)
  movel([0.261420, -1.166933, -2.691745, -0.853711, 1.570796, 1.832217],accel_mss,speed_ms,0,blend_radius_m)
  movel([0.264066, -1.163130, -2.693415, -0.855844, 1.570796, 1.834862],accel_mss,speed_ms,0,blend_radius_m)
  movel([0.267036, -1.159707, -2.694905, -0.857777, 1.570796, 1.837832],accel_mss,speed_ms,0,blend_radius_m)
  movel([0.270280, -1.156643, -2.696229, -0.859518, 1.570796, 1.841076],accel_mss,speed_ms,0,blend_radius_m)
  movel([0.273744, -1.153912, -2.697400, -0.861077, 1.570796, 1.844541],accel_mss,speed_ms,0,blend_radius_m)
  movel([0.277383, -1.151488, -2.698434, -0.862467, 1.570796, 1.848179],accel_mss,speed_ms,0,blend_radius_m)
  movel([0.281137, -1.149344, -2.699343, -0.863702, 1.570796, 1.851933],accel_mss,speed_ms,0,blend_radius_m)
  movel([0.284960, -1.147449, -2.700143, -0.864797, 1.570796, 1.855756],accel_mss,speed_ms,0,blend_radius_m)
  movel([0.288796, -1.145776, -2.700846, -0.865767, 1.570796, 1.859592],accel_mss,speed_ms,0,blend_radius_m)
  movel([0.295860, -1.143294, -2.701884, -0.867211, 1.570796, 1.866656],accel_mss,speed_ms,0,blend_radius_m)
  movel([0.301777, -1.141931, -2.702452, -0.868006, 1.570796, 1.872573],accel_mss,speed_ms,0,blend_radius_m)
  movel([0.306468, -1.141416, -2.702665, -0.868307, 1.570796, 1.877264],accel_mss,speed_ms,0,blend_radius_m)
  movel([0.309865, -1.141460, -2.702647, -0.868282, 1.570796, 1.880661],accel_mss,speed_ms,0,blend_radius_m)
  movel([0.314427, -1.142309, -2.702294, -0.867786, 1.570796, 1.885223],accel_mss,speed_ms,0,blend_radius_m)
  movel([0.318299, -1.143981, -2.701597, -0.866811, 1.570796, 1.889095],accel_mss,speed_ms,0,blend_radius_m)
  movel([0.321475, -1.146401, -2.700584, -0.865404, 1.570796, 1.892272],accel_mss,speed_ms,0,blend_radius_m)
  movel([0.323949, -1.149490, -2.699281, -0.863618, 1.570796, 1.894746],accel_mss,speed_ms,0,blend_radius_m)
  movel([0.325716, -1.153164, -2.697720, -0.861505, 1.570796, 1.896512],accel_mss,speed_ms,0,blend_radius_m)
  movel([0.326777, -1.157341, -2.695928, -0.859120, 1.570796, 1.897573],accel_mss,speed_ms,0,blend_radius_m)
  movel([0.327132, -1.161949, -2.693930, -0.856510, 1.570796, 1.897929],accel_mss,speed_ms,0,blend_radius_m)
  movel([0.326787, -1.166904, -2.691758, -0.853727, 1.570796, 1.897583],accel_mss,speed_ms,0,blend_radius_m)
  movel([0.325876, -1.171601, -2.689675, -0.851112, 1.570796, 1.896672],accel_mss,speed_ms,0,blend_radius_m)
  movel([0.324622, -1.176358, -2.687543, -0.848488, 1.570796, 1.895419],accel_mss,speed_ms,0,blend_radius_m)
  movel([0.323338, -1.181031, -2.685425, -0.845933, 1.570796, 1.894134],accel_mss,speed_ms,0,blend_radius_m)
  movel([0.322340, -1.185483, -2.683385, -0.843521, 1.570796, 1.893136],accel_mss,speed_ms,0,blend_radius_m)
  movel([0.321932, -1.189573, -2.681493, -0.841323, 1.570796, 1.892729],accel_mss,speed_ms,0,blend_radius_m)
  movel([0.322044, -1.191442, -2.680622, -0.840325, 1.570796, 1.892840],accel_mss,speed_ms,0,blend_radius_m)
  movel([0.322416, -1.193176, -2.679811, -0.839403, 1.570796, 1.893212],accel_mss,speed_ms,0,blend_radius_m)
  movel([0.323087, -1.194753, -2.679070, -0.838566, 1.570796, 1.893883],accel_mss,speed_ms,0,blend_radius_m)
  movel([0.324093, -1.196164, -2.678405, -0.837820, 1.570796, 1.894889],accel_mss,speed_ms,0,blend_radius_m)
  movel([0.325466, -1.197391, -2.677825, -0.837173, 1.570796, 1.896263],accel_mss,speed_ms,0,blend_radius_m)
  movel([0.327251, -1.198421, -2.677337, -0.836631, 1.570796, 1.898047],accel_mss,speed_ms,0,blend_radius_m)
  movel([0.329089, -1.198965, -2.677078, -0.836345, 1.570796, 1.899886],accel_mss,speed_ms,0,blend_radius_m)
  movel([0.330960, -1.198964, -2.677079, -0.836346, 1.570796, 1.901756],accel_mss,speed_ms,0,blend_radius_m)
  movel([0.332825, -1.198495, -2.677302, -0.836592, 1.570796, 1.903622],accel_mss,speed_ms,0,blend_radius_m)
  movel([0.334640, -1.197627, -2.677713, -0.837049, 1.570796, 1.905437],accel_mss,speed_ms,0,blend_radius_m)
  movel([0.336368, -1.196433, -2.678278, -0.837678, 1.570796, 1.907164],accel_mss,speed_ms,0,blend_radius_m)
  movel([0.337961, -1.194988, -2.678959, -0.838442, 1.570796, 1.908757],accel_mss,speed_ms,0,blend_radius_m)
  movel([0.339377, -1.193359, -2.679725, -0.839305, 1.570796, 1.910173],accel_mss,speed_ms,0,blend_radius_m)
  movel([0.340570, -1.191622, -2.680538, -0.840229, 1.570796, 1.911367],accel_mss,speed_ms,0,blend_radius_m)
  movel([0.341498, -1.189852, -2.681363, -0.841174, 1.570796, 1.912294],accel_mss,speed_ms,0,blend_radius_m)
  movel([0.342112, -1.188122, -2.682166, -0.842101, 1.570796, 1.912908],accel_mss,speed_ms,0,blend_radius_m)
  movel([0.342365, -1.186512, -2.682911, -0.842966, 1.570796, 1.913161],accel_mss,speed_ms,0,blend_radius_m)
  movel([0.342210, -1.185093, -2.683565, -0.843731, 1.570796, 1.913007],accel_mss,speed_ms,0,blend_radius_m)
  movel([0.341597, -1.183952, -2.684089, -0.844348, 1.570796, 1.912393],accel_mss,speed_ms,0,blend_radius_m)
  movel([0.340482, -1.183164, -2.684450, -0.844775, 1.570796, 1.911278],accel_mss,speed_ms,0,blend_radius_m)
  movel([0.338820, -1.182807, -2.684614, -0.844969, 1.570796, 1.909616],accel_mss,speed_ms,0,blend_radius_m)
  movel([0.336560, -1.182965, -2.684541, -0.844882, 1.570796, 1.907356],accel_mss,speed_ms,0,blend_radius_m)
  movel([0.337123, -1.184067, -2.684036, -0.844286, 1.570796, 1.907919],accel_mss,speed_ms,0,blend_radius_m)
  movel([0.337304, -1.185232, -2.683501, -0.843656, 1.570796, 1.908100],accel_mss,speed_ms,0,blend_radius_m)
  movel([0.337125, -1.186413, -2.682956, -0.843019, 1.570796, 1.907921],accel_mss,speed_ms,0,blend_radius_m)
  movel([0.336607, -1.187558, -2.682427, -0.842404, 1.570796, 1.907403],accel_mss,speed_ms,0,blend_radius_m)
  movel([0.335771, -1.188629, -2.681931, -0.841829, 1.570796, 1.906567],accel_mss,speed_ms,0,blend_radius_m)
  movel([0.334643, -1.189572, -2.681493, -0.841324, 1.570796, 1.905439],accel_mss,speed_ms,0,blend_radius_m)
  movel([0.333235, -1.190342, -2.681135, -0.840912, 1.570796, 1.904032],accel_mss,speed_ms,0,blend_radius_m)
  movel([0.331573, -1.190901, -2.680874, -0.840614, 1.570796, 1.902369],accel_mss,speed_ms,0,blend_radius_m)
  movel([0.328913, -1.191215, -2.680728, -0.840446, 1.570796, 1.899710],accel_mss,speed_ms,0,blend_radius_m)
  movel([0.326905, -1.190765, -2.680938, -0.840686, 1.570796, 1.897701],accel_mss,speed_ms,0,blend_radius_m)
  movel([0.325508, -1.189643, -2.681460, -0.841286, 1.570796, 1.896305],accel_mss,speed_ms,0,blend_radius_m)
  movel([0.324691, -1.187955, -2.682243, -0.842190, 1.570796, 1.895487],accel_mss,speed_ms,0,blend_radius_m)
  movel([0.324419, -1.185788, -2.683245, -0.843356, 1.570796, 1.895215],accel_mss,speed_ms,0,blend_radius_m)
  movel([0.324661, -1.183244, -2.684414, -0.844732, 1.570796, 1.895457],accel_mss,speed_ms,0,blend_radius_m)
  movel([0.325387, -1.180414, -2.685706, -0.846269, 1.570796, 1.896183],accel_mss,speed_ms,0,blend_radius_m)
  movel([0.326563, -1.177404, -2.687071, -0.847914, 1.570796, 1.897359],accel_mss,speed_ms,0,blend_radius_m)
  movel([0.328164, -1.174309, -2.688464, -0.849616, 1.570796, 1.898961],accel_mss,speed_ms,0,blend_radius_m)
  movel([0.330154, -1.171235, -2.689838, -0.851315, 1.570796, 1.900950],accel_mss,speed_ms,0,blend_radius_m)
  movel([0.332497, -1.168288, -2.691147, -0.852954, 1.570796, 1.903293],accel_mss,speed_ms,0,blend_radius_m)
  movel([0.335158, -1.165578, -2.692342, -0.854469, 1.570796, 1.905955],accel_mss,speed_ms,0,blend_radius_m)
  movel([0.338102, -1.163218, -2.693377, -0.855795, 1.570796, 1.908899],accel_mss,speed_ms,0,blend_radius_m)
  movel([0.341285, -1.161318, -2.694205, -0.856866, 1.570796, 1.912081],accel_mss,speed_ms,0,blend_radius_m)
  movel([0.344668, -1.159993, -2.694781, -0.857615, 1.570796, 1.915465],accel_mss,speed_ms,0,blend_radius_m)
  movel([0.348203, -1.159360, -2.695055, -0.857974, 1.570796, 1.918999],accel_mss,speed_ms,0,blend_radius_m)
  movel([0.350586, -1.159329, -2.695069, -0.857992, 1.570796, 1.921383],accel_mss,speed_ms,0,blend_radius_m)
  movel([0.352804, -1.159566, -2.694966, -0.857857, 1.570796, 1.923600],accel_mss,speed_ms,0,blend_radius_m)
  movel([0.354842, -1.160066, -2.694749, -0.857574, 1.570796, 1.925638],accel_mss,speed_ms,0,blend_radius_m)
  movel([0.356684, -1.160814, -2.694424, -0.857151, 1.570796, 1.927481],accel_mss,speed_ms,0,blend_radius_m)
  movel([0.358322, -1.161801, -2.693995, -0.856593, 1.570796, 1.929118],accel_mss,speed_ms,0,blend_radius_m)
  movel([0.359744, -1.163015, -2.693465, -0.855909, 1.570796, 1.930540],accel_mss,speed_ms,0,blend_radius_m)
  movel([0.360932, -1.164442, -2.692841, -0.855107, 1.570796, 1.931728],accel_mss,speed_ms,0,blend_radius_m)
  movel([0.361881, -1.166070, -2.692125, -0.854193, 1.570796, 1.932677],accel_mss,speed_ms,0,blend_radius_m)
  movel([0.362573, -1.167889, -2.691323, -0.853177, 1.570796, 1.933369],accel_mss,speed_ms,0,blend_radius_m)
  movel([0.363005, -1.169885, -2.690439, -0.852065, 1.570796, 1.933801],accel_mss,speed_ms,0,blend_radius_m)
  movel([0.363161, -1.172046, -2.689477, -0.850866, 1.570796, 1.933958],accel_mss,speed_ms,0,blend_radius_m)
  movel([0.363038, -1.174357, -2.688443, -0.849589, 1.570796, 1.933834],accel_mss,speed_ms,0,blend_radius_m)
  movel([0.362615, -1.176812, -2.687338, -0.848239, 1.570796, 1.933412],accel_mss,speed_ms,0,blend_radius_m)
  movel([0.361891, -1.179393, -2.686170, -0.846826, 1.570796, 1.932687],accel_mss,speed_ms,0,blend_radius_m)
  movel([0.360854, -1.182091, -2.684941, -0.845357, 1.570796, 1.931651],accel_mss,speed_ms,0,blend_radius_m)
  movel([0.359494, -1.184896, -2.683655, -0.843838, 1.570796, 1.930290],accel_mss,speed_ms,0,blend_radius_m)
  movel([0.357637, -1.187617, -2.682400, -0.842372, 1.570796, 1.928434],accel_mss,speed_ms,0,blend_radius_m)
  movel([0.355252, -1.190441, -2.681089, -0.840859, 1.570796, 1.926048],accel_mss,speed_ms,0,blend_radius_m)
  movel([0.353108, -1.192822, -2.679976, -0.839590, 1.570796, 1.923904],accel_mss,speed_ms,0,blend_radius_m)
  movel([0.351972, -1.194223, -2.679319, -0.838847, 1.570796, 1.922769],accel_mss,speed_ms,0,blend_radius_m)
  movel([0.351833, -1.195360, -2.678784, -0.838245, 1.570796, 1.922630],accel_mss,speed_ms,0,blend_radius_m)
  movel([0.351996, -1.197047, -2.677988, -0.837354, 1.570796, 1.922793],accel_mss,speed_ms,0,blend_radius_m)
  movel([0.352182, -1.198900, -2.677109, -0.836379, 1.570796, 1.922978],accel_mss,speed_ms,0,blend_radius_m)
  movel([0.352109, -1.200540, -2.676329, -0.835520, 1.570796, 1.922905],accel_mss,speed_ms,0,blend_radius_m)
  movel([0.351459, -1.202877, -2.675212, -0.834301, 1.570796, 1.922255],accel_mss,speed_ms,0,blend_radius_m)
  movel([0.350520, -1.205119, -2.674134, -0.833136, 1.570796, 1.921316],accel_mss,speed_ms,0,blend_radius_m)
  movel([0.349328, -1.207258, -2.673100, -0.832031, 1.570796, 1.920124],accel_mss,speed_ms,0,blend_radius_m)
  movel([0.347916, -1.209272, -2.672123, -0.830994, 1.570796, 1.918713],accel_mss,speed_ms,0,blend_radius_m)
  movel([0.346315, -1.211151, -2.671206, -0.830031, 1.570796, 1.917111],accel_mss,speed_ms,0,blend_radius_m)
  movel([0.344553, -1.212881, -2.670360, -0.829148, 1.570796, 1.915349],accel_mss,speed_ms,0,blend_radius_m)
  movel([0.342665, -1.214444, -2.669591, -0.828353, 1.570796, 1.913461],accel_mss,speed_ms,0,blend_radius_m)
  movel([0.340680, -1.215832, -2.668907, -0.827650, 1.570796, 1.911476],accel_mss,speed_ms,0,blend_radius_m)
  movel([0.338624, -1.217027, -2.668316, -0.827046, 1.570796, 1.909420],accel_mss,speed_ms,0,blend_radius_m)
  movel([0.336533, -1.218016, -2.667826, -0.826547, 1.570796, 1.907329],accel_mss,speed_ms,0,blend_radius_m)
  movel([0.334430, -1.218783, -2.667445, -0.826162, 1.570796, 1.905226],accel_mss,speed_ms,0,blend_radius_m)
  speed_ms = 0.003
  movel([0.334430, -1.211558, -2.663890, -0.836941, 1.570796, 1.905226],accel_mss,speed_ms,0,blend_radius_m)
  speed_ms = 1.000
  movel([0.334430, -1.184074, -2.649412, -0.878903, 1.570796, 1.905226],accel_mss,speed_ms,0,blend_radius_m)
  #M_RunCode9
  movel([0.342398, -1.190482, -2.646347, -0.875560, 1.570796, 1.913195],accel_mss,speed_ms,0,blend_radius_m)
  #M_RunCode3
  movel([0.342398, -1.217908, -2.660741, -0.833740, 1.570796, 1.913195],accel_mss,speed_ms,0,blend_radius_m)
  speed_ms = 0.003
  movel([0.342398, -1.225114, -2.664274, -0.823001, 1.570796, 1.913195],accel_mss,speed_ms,0,blend_radius_m)
  speed_ms = 0.007
  movel([0.343849, -1.223656, -2.665008, -0.823725, 1.570796, 1.914646],accel_mss,speed_ms,0,blend_radius_m)
  movel([0.347050, -1.220946, -2.666366, -0.825076, 1.570796, 1.917846],accel_mss,speed_ms,0,blend_radius_m)
  movel([0.350088, -1.218214, -2.667727, -0.826448, 1.570796, 1.920884],accel_mss,speed_ms,0,blend_radius_m)
  movel([0.351332, -1.216727, -2.668464, -0.827197, 1.570796, 1.922128],accel_mss,speed_ms,0,blend_radius_m)
  movel([0.352284, -1.215096, -2.669270, -0.828023, 1.570796, 1.923080],accel_mss,speed_ms,0,blend_radius_m)
  movel([0.351928, -1.216289, -2.668681, -0.827419, 1.570796, 1.922724],accel_mss,speed_ms,0,blend_radius_m)
  movel([0.350906, -1.218471, -2.667600, -0.826319, 1.570796, 1.921703],accel_mss,speed_ms,0,blend_radius_m)
  movel([0.349568, -1.220411, -2.666634, -0.825345, 1.570796, 1.920365],accel_mss,speed_ms,0,blend_radius_m)
  movel([0.348005, -1.222194, -2.665742, -0.824453, 1.570796, 1.918801],accel_mss,speed_ms,0,blend_radius_m)
  movel([0.346319, -1.223888, -2.664891, -0.823610, 1.570796, 1.917115],accel_mss,speed_ms,0,blend_radius_m)
  movel([0.342958, -1.227317, -2.663160, -0.821913, 1.570796, 1.913754],accel_mss,speed_ms,0,blend_radius_m)
  movel([0.341482, -1.229198, -2.662203, -0.820987, 1.570796, 1.912278],accel_mss,speed_ms,0,blend_radius_m)
  movel([0.340271, -1.231284, -2.661139, -0.819966, 1.570796, 1.911067],accel_mss,speed_ms,0,blend_radius_m)
  movel([0.339299, -1.233663, -2.659918, -0.818807, 1.570796, 1.910095],accel_mss,speed_ms,0,blend_radius_m)
  movel([0.338886, -1.234925, -2.659268, -0.818195, 1.570796, 1.909682],accel_mss,speed_ms,0,blend_radius_m)
  movel([0.338807, -1.235625, -2.658907, -0.817857, 1.570796, 1.909603],accel_mss,speed_ms,0,blend_radius_m)
  movel([0.339712, -1.235790, -2.658822, -0.817777, 1.570796, 1.910508],accel_mss,speed_ms,0,blend_radius_m)
  movel([0.340424, -1.235971, -2.658728, -0.817689, 1.570796, 1.911220],accel_mss,speed_ms,0,blend_radius_m)
  movel([0.341025, -1.236338, -2.658539, -0.817513, 1.570796, 1.911822],accel_mss,speed_ms,0,blend_radius_m)
  movel([0.341858, -1.237439, -2.657968, -0.816982, 1.570796, 1.912655],accel_mss,speed_ms,0,blend_radius_m)
  movel([0.342225, -1.238495, -2.657420, -0.816474, 1.570796, 1.913021],accel_mss,speed_ms,0,blend_radius_m)
  movel([0.342211, -1.239538, -2.656877, -0.815974, 1.570796, 1.913008],accel_mss,speed_ms,0,blend_radius_m)
  movel([0.341912, -1.240600, -2.656322, -0.815467, 1.570796, 1.912708],accel_mss,speed_ms,0,blend_radius_m)
  movel([0.340799, -1.242907, -2.655114, -0.814368, 1.570796, 1.911596],accel_mss,speed_ms,0,blend_radius_m)
  movel([0.339590, -1.245676, -2.653655, -0.813058, 1.570796, 1.910386],accel_mss,speed_ms,0,blend_radius_m)
  movel([0.338526, -1.249345, -2.651708, -0.811336, 1.570796, 1.909322],accel_mss,speed_ms,0,blend_radius_m)
  movel([0.337606, -1.252957, -2.649775, -0.809657, 1.570796, 1.908402],accel_mss,speed_ms,0,blend_radius_m)
  movel([0.336534, -1.256574, -2.647824, -0.807990, 1.570796, 1.907331],accel_mss,speed_ms,0,blend_radius_m)
  movel([0.335031, -1.260245, -2.645828, -0.806316, 1.570796, 1.905827],accel_mss,speed_ms,0,blend_radius_m)
  movel([0.333945, -1.262228, -2.644743, -0.805418, 1.570796, 1.904741],accel_mss,speed_ms,0,blend_radius_m)
  movel([0.332683, -1.264172, -2.643674, -0.804543, 1.570796, 1.903479],accel_mss,speed_ms,0,blend_radius_m)
  movel([0.329831, -1.267949, -2.641585, -0.802855, 1.570796, 1.900627],accel_mss,speed_ms,0,blend_radius_m)
  movel([0.326847, -1.271609, -2.639544, -0.801236, 1.570796, 1.897643],accel_mss,speed_ms,0,blend_radius_m)
  movel([0.324113, -1.275171, -2.637541, -0.799676, 1.570796, 1.894909],accel_mss,speed_ms,0,blend_radius_m)
  movel([0.320194, -1.281214, -2.634108, -0.797067, 1.570796, 1.890991],accel_mss,speed_ms,0,blend_radius_m)
  movel([0.318581, -1.283801, -2.632624, -0.795964, 1.570796, 1.889377],accel_mss,speed_ms,0,blend_radius_m)
  movel([0.316934, -1.286205, -2.631237, -0.794946, 1.570796, 1.887730],accel_mss,speed_ms,0,blend_radius_m)
  movel([0.315062, -1.288497, -2.629909, -0.793983, 1.570796, 1.885858],accel_mss,speed_ms,0,blend_radius_m)
  movel([0.312769, -1.290758, -2.628592, -0.793039, 1.570796, 1.883565],accel_mss,speed_ms,0,blend_radius_m)
  movel([0.309864, -1.293062, -2.627243, -0.792085, 1.570796, 1.880660],accel_mss,speed_ms,0,blend_radius_m)
  movel([0.306156, -1.295486, -2.625816, -0.791087, 1.570796, 1.876952],accel_mss,speed_ms,0,blend_radius_m)
  movel([0.303064, -1.297203, -2.624801, -0.790385, 1.570796, 1.873860],accel_mss,speed_ms,0,blend_radius_m)
  movel([0.300187, -1.298517, -2.624021, -0.789850, 1.570796, 1.870983],accel_mss,speed_ms,0,blend_radius_m)
  movel([0.297508, -1.299456, -2.623463, -0.789470, 1.570796, 1.868304],accel_mss,speed_ms,0,blend_radius_m)
  movel([0.295020, -1.300045, -2.623112, -0.789232, 1.570796, 1.865816],accel_mss,speed_ms,0,blend_radius_m)
  movel([0.292716, -1.300301, -2.622960, -0.789128, 1.570796, 1.863512],accel_mss,speed_ms,0,blend_radius_m)
  movel([0.290588, -1.300249, -2.622991, -0.789149, 1.570796, 1.861384],accel_mss,speed_ms,0,blend_radius_m)
  movel([0.288623, -1.299910, -2.623193, -0.789286, 1.570796, 1.859419],accel_mss,speed_ms,0,blend_radius_m)
  movel([0.286816, -1.299304, -2.623554, -0.789532, 1.570796, 1.857612],accel_mss,speed_ms,0,blend_radius_m)
  movel([0.285163, -1.298453, -2.624059, -0.789876, 1.570796, 1.855959],accel_mss,speed_ms,0,blend_radius_m)
  movel([0.283653, -1.297380, -2.624696, -0.790313, 1.570796, 1.854449],accel_mss,speed_ms,0,blend_radius_m)
  movel([0.281044, -1.294639, -2.626315, -0.791435, 1.570796, 1.851840],accel_mss,speed_ms,0,blend_radius_m)
  movel([0.278941, -1.291244, -2.628308, -0.792837, 1.570796, 1.849737],accel_mss,speed_ms,0,blend_radius_m)
  movel([0.277300, -1.287356, -2.630571, -0.794462, 1.570796, 1.848097],accel_mss,speed_ms,0,blend_radius_m)
  movel([0.276212, -1.283361, -2.632877, -0.796151, 1.570796, 1.847008],accel_mss,speed_ms,0,blend_radius_m)
  movel([0.274935, -1.278134, -2.635864, -0.798391, 1.570796, 1.845732],accel_mss,speed_ms,0,blend_radius_m)
  movel([0.273199, -1.272511, -2.639038, -0.800840, 1.570796, 1.843995],accel_mss,speed_ms,0,blend_radius_m)
  movel([0.272072, -1.269815, -2.640547, -0.802027, 1.570796, 1.842868],accel_mss,speed_ms,0,blend_radius_m)
  movel([0.270726, -1.267346, -2.641920, -0.803123, 1.570796, 1.841522],accel_mss,speed_ms,0,blend_radius_m)
  movel([0.269127, -1.265217, -2.643098, -0.804074, 1.570796, 1.839923],accel_mss,speed_ms,0,blend_radius_m)
  movel([0.267242, -1.263536, -2.644025, -0.804829, 1.570796, 1.838038],accel_mss,speed_ms,0,blend_radius_m)
  movel([0.265038, -1.262417, -2.644639, -0.805333, 1.570796, 1.835835],accel_mss,speed_ms,0,blend_radius_m)
  movel([0.262488, -1.261972, -2.644883, -0.805534, 1.570796, 1.833285],accel_mss,speed_ms,0,blend_radius_m)
  movel([0.261071, -1.262040, -2.644846, -0.805503, 1.570796, 1.831868],accel_mss,speed_ms,0,blend_radius_m)
  movel([0.259560, -1.262315, -2.644695, -0.805379, 1.570796, 1.830356],accel_mss,speed_ms,0,blend_radius_m)
  movel([0.257946, -1.262816, -2.644420, -0.805153, 1.570796, 1.828742],accel_mss,speed_ms,0,blend_radius_m)
  movel([0.256232, -1.263549, -2.644017, -0.804822, 1.570796, 1.827028],accel_mss,speed_ms,0,blend_radius_m)
  movel([0.254410, -1.264533, -2.643475, -0.804380, 1.570796, 1.825207],accel_mss,speed_ms,0,blend_radius_m)
  movel([0.252483, -1.265776, -2.642789, -0.803824, 1.570796, 1.823279],accel_mss,speed_ms,0,blend_radius_m)
  movel([0.248294, -1.269094, -2.640948, -0.802346, 1.570796, 1.819091],accel_mss,speed_ms,0,blend_radius_m)
  movel([0.246565, -1.270999, -2.639885, -0.801505, 1.570796, 1.817361],accel_mss,speed_ms,0,blend_radius_m)
  movel([0.245072, -1.273098, -2.638709, -0.800582, 1.570796, 1.815868],accel_mss,speed_ms,0,blend_radius_m)
  movel([0.243850, -1.275378, -2.637424, -0.799586, 1.570796, 1.814646],accel_mss,speed_ms,0,blend_radius_m)
  movel([0.242932, -1.277824, -2.636040, -0.798525, 1.570796, 1.813729],accel_mss,speed_ms,0,blend_radius_m)
  movel([0.245868, -1.276117, -2.637007, -0.799265, 1.570796, 1.816664],accel_mss,speed_ms,0,blend_radius_m)
  movel([0.248749, -1.274733, -2.637788, -0.799867, 1.570796, 1.819545],accel_mss,speed_ms,0,blend_radius_m)
  movel([0.251553, -1.273667, -2.638389, -0.800333, 1.570796, 1.822349],accel_mss,speed_ms,0,blend_radius_m)
  movel([0.254263, -1.272918, -2.638810, -0.800661, 1.570796, 1.825059],accel_mss,speed_ms,0,blend_radius_m)
  movel([0.256853, -1.272482, -2.639054, -0.800852, 1.570796, 1.827649],accel_mss,speed_ms,0,blend_radius_m)
  movel([0.259307, -1.272351, -2.639128, -0.800910, 1.570796, 1.830104],accel_mss,speed_ms,0,blend_radius_m)
  movel([0.261601, -1.272527, -2.639029, -0.800833, 1.570796, 1.832397],accel_mss,speed_ms,0,blend_radius_m)
  movel([0.263716, -1.272997, -2.638766, -0.800626, 1.570796, 1.834512],accel_mss,speed_ms,0,blend_radius_m)
  movel([0.265631, -1.273761, -2.638336, -0.800292, 1.570796, 1.836427],accel_mss,speed_ms,0,blend_radius_m)
  movel([0.267332, -1.274806, -2.637747, -0.799835, 1.570796, 1.838128],accel_mss,speed_ms,0,blend_radius_m)
  movel([0.268797, -1.276126, -2.637002, -0.799261, 1.570796, 1.839593],accel_mss,speed_ms,0,blend_radius_m)
  movel([0.270009, -1.277714, -2.636102, -0.798573, 1.570796, 1.840805],accel_mss,speed_ms,0,blend_radius_m)
  movel([0.270950, -1.279560, -2.635052, -0.797777, 1.570796, 1.841746],accel_mss,speed_ms,0,blend_radius_m)
  movel([0.271604, -1.281657, -2.633854, -0.796877, 1.570796, 1.842401],accel_mss,speed_ms,0,blend_radius_m)
  movel([0.271955, -1.283995, -2.632513, -0.795882, 1.570796, 1.842752],accel_mss,speed_ms,0,blend_radius_m)
  movel([0.271991, -1.286565, -2.631029, -0.794795, 1.570796, 1.842788],accel_mss,speed_ms,0,blend_radius_m)
  movel([0.271770, -1.288784, -2.629742, -0.793863, 1.570796, 1.842566],accel_mss,speed_ms,0,blend_radius_m)
  movel([0.271333, -1.290994, -2.628454, -0.792941, 1.570796, 1.842129],accel_mss,speed_ms,0,blend_radius_m)
  movel([0.270694, -1.293186, -2.627170, -0.792033, 1.570796, 1.841491],accel_mss,speed_ms,0,blend_radius_m)
  movel([0.269872, -1.295347, -2.625898, -0.791144, 1.570796, 1.840669],accel_mss,speed_ms,0,blend_radius_m)
  movel([0.267730, -1.299550, -2.623407, -0.789432, 1.570796, 1.838526],accel_mss,speed_ms,0,blend_radius_m)
  movel([0.265020, -1.303531, -2.621027, -0.787831, 1.570796, 1.835816],accel_mss,speed_ms,0,blend_radius_m)
  movel([0.261857, -1.307222, -2.618801, -0.786366, 1.570796, 1.832654],accel_mss,speed_ms,0,blend_radius_m)
  movel([0.258353, -1.310556, -2.616776, -0.785057, 1.570796, 1.829149],accel_mss,speed_ms,0,blend_radius_m)
  movel([0.254607, -1.313472, -2.614993, -0.783925, 1.570796, 1.825404],accel_mss,speed_ms,0,blend_radius_m)
  movel([0.250727, -1.315901, -2.613498, -0.782990, 1.570796, 1.821523],accel_mss,speed_ms,0,blend_radius_m)
  movel([0.246810, -1.317781, -2.612337, -0.782271, 1.570796, 1.817607],accel_mss,speed_ms,0,blend_radius_m)
  movel([0.242960, -1.319047, -2.611551, -0.781790, 1.570796, 1.813756],accel_mss,speed_ms,0,blend_radius_m)
  movel([0.239272, -1.319630, -2.611189, -0.781570, 1.570796, 1.810068],accel_mss,speed_ms,0,blend_radius_m)
  movel([0.237519, -1.319646, -2.611180, -0.781564, 1.570796, 1.808315],accel_mss,speed_ms,0,blend_radius_m)
  movel([0.235843, -1.319461, -2.611294, -0.781633, 1.570796, 1.806640],accel_mss,speed_ms,0,blend_radius_m)
  movel([0.234256, -1.319073, -2.611535, -0.781780, 1.570796, 1.805053],accel_mss,speed_ms,0,blend_radius_m)
  movel([0.232773, -1.318466, -2.611912, -0.782011, 1.570796, 1.803569],accel_mss,speed_ms,0,blend_radius_m)
  movel([0.231401, -1.317633, -2.612428, -0.782328, 1.570796, 1.802198],accel_mss,speed_ms,0,blend_radius_m)
  movel([0.230159, -1.316564, -2.613089, -0.782736, 1.570796, 1.800955],accel_mss,speed_ms,0,blend_radius_m)
  movel([0.229057, -1.315248, -2.613901, -0.783240, 1.570796, 1.799853],accel_mss,speed_ms,0,blend_radius_m)
  movel([0.228109, -1.313673, -2.614869, -0.783847, 1.570796, 1.798905],accel_mss,speed_ms,0,blend_radius_m)
  movel([0.227326, -1.311827, -2.616000, -0.784562, 1.570796, 1.798123],accel_mss,speed_ms,0,blend_radius_m)
  movel([0.226725, -1.309699, -2.617298, -0.785392, 1.570796, 1.797522],accel_mss,speed_ms,0,blend_radius_m)
  movel([0.226563, -1.307778, -2.618465, -0.786146, 1.570796, 1.797360],accel_mss,speed_ms,0,blend_radius_m)
  movel([0.226646, -1.302193, -2.621829, -0.788367, 1.570796, 1.797442],accel_mss,speed_ms,0,blend_radius_m)
  movel([0.227050, -1.298096, -2.624271, -0.790022, 1.570796, 1.797846],accel_mss,speed_ms,0,blend_radius_m)
  movel([0.227842, -1.293163, -2.627183, -0.792043, 1.570796, 1.798638],accel_mss,speed_ms,0,blend_radius_m)
  movel([0.229147, -1.287409, -2.630541, -0.794440, 1.570796, 1.799943],accel_mss,speed_ms,0,blend_radius_m)
  movel([0.231078, -1.280852, -2.634315, -0.797222, 1.570796, 1.801875],accel_mss,speed_ms,0,blend_radius_m)
  movel([0.232808, -1.276165, -2.636980, -0.799244, 1.570796, 1.803605],accel_mss,speed_ms,0,blend_radius_m)
  movel([0.234755, -1.271863, -2.639402, -0.801124, 1.570796, 1.805551],accel_mss,speed_ms,0,blend_radius_m)
  movel([0.236872, -1.267938, -2.641592, -0.802860, 1.570796, 1.807668],accel_mss,speed_ms,0,blend_radius_m)
  movel([0.239118, -1.264382, -2.643559, -0.804448, 1.570796, 1.809914],accel_mss,speed_ms,0,blend_radius_m)
  movel([0.241446, -1.261188, -2.645313, -0.805888, 1.570796, 1.812242],accel_mss,speed_ms,0,blend_radius_m)
  movel([0.243811, -1.258344, -2.646864, -0.807181, 1.570796, 1.814608],accel_mss,speed_ms,0,blend_radius_m)
  movel([0.246168, -1.255837, -2.648223, -0.808329, 1.570796, 1.816964],accel_mss,speed_ms,0,blend_radius_m)
  movel([0.248471, -1.253660, -2.649397, -0.809332, 1.570796, 1.819267],accel_mss,speed_ms,0,blend_radius_m)
  movel([0.252723, -1.250231, -2.651235, -0.810923, 1.570796, 1.823520],accel_mss,speed_ms,0,blend_radius_m)
  movel([0.256206, -1.247947, -2.652452, -0.811990, 1.570796, 1.827002],accel_mss,speed_ms,0,blend_radius_m)
  movel([0.258552, -1.246678, -2.653125, -0.812586, 1.570796, 1.829348],accel_mss,speed_ms,0,blend_radius_m)
  movel([0.259412, -1.246286, -2.653332, -0.812771, 1.570796, 1.830209],accel_mss,speed_ms,0,blend_radius_m)
  movel([0.263427, -1.244750, -2.654144, -0.813495, 1.570796, 1.834223],accel_mss,speed_ms,0,blend_radius_m)
